(* IEC 61131-3 sources: daoli-st-library/DL_Motion (part 18) *)

(* ---- FB_DL_StackingAlignCtrl.st ---- *)
//==============================================================================
// 功能块：FB_DL_StackingAlignCtrl ｜ 中文名称：叠片对位纠偏控制
// 所属子库：DL_Motion ｜ 版本：v1.0.0 ｜ 兼容：CODESYS V3.5+ / TwinCAT 3 / 汇川 InoProShop
// 功能描述：叠片机 CCD 对位纠偏量的解算件。输入像素偏差与角度偏差，经「像素→机械」
//           标定矩阵的逆映射得机械纠偏量（mm / mrad），输出双轴纠偏指令、超差 NG 与
//           行程限幅标志。标定矩阵求逆委托 FC_DL_Affine2DInvert（组合调用，不复制
//           低层实现）；矩阵奇异时沿用上次有效逆矩阵并置 bMatrixFallback，无历史有效
//           值时判故障。本件只解算纠偏量，不定义轴状态、不发运动指令——轴状态与运动
//           指令的唯一属主是运动层（T1-6 纪律），本件仅输出「允许上层下发纠偏」的
//           bReady 许可位。
// 开源溯源 (Origin)：道莅原创实现（参考 公开工程惯例 分类与参数域）
// 单位表：像素偏差[像素] / 纠偏量[mm] / 角度偏差与角度纠偏量[mrad] / 标定矩阵线性块
//         [mm 每像素] / 标定矩阵平移列[mm] / 行程门限[mm] / 超差门限[mm 或 mrad] /
//         行列式[无量纲]
// 错误码表：16#0004_01EB 信息级（纠偏量被行程限幅，bClamped 置位，限幅后值不得当作
//           正常纠偏量计数，须 HMI 可辨，不置 bError）/ 16#0004_01EC 信息级（标定矩阵
//           退化不可逆，沿用上次有效逆矩阵，bMatrixFallback 置位，不置 bError）/
//           16#0004_030C 故障级（标定矩阵非法/不可逆且无历史有效值，置 bError，纠偏量
//           回零）/ 16#0004_030D 故障级（输入非有限或纠偏解算溢出，置 bError，纠偏量
//           回零）/ 16#0004_030E 故障级兜底（状态机落 ELSE 非法状态，置 bError，纠偏量
//           回零）。码位 16#0004 段，信息带 01xx、故障带 03xx，不越段不挪用预留槽。
// 状态机：E_DL_StackAlignState（eIdle=0 失能/待机 / eAlign=10 正常纠偏解算 /
//           eLimited=20 行程限幅生效 / eCamLost=30 相机无效不纠偏 / eFault=99 故障
//           兜底），CASE 含 ELSE 兜底，ELSE 置 030E 且纠偏量回零 bValid := FALSE。
// 边界行为：① 标定矩阵经 FC_DL_Affine2DInvert 求逆（每拍无条件调用恰好一次）；奇异
//           时若有历史有效逆矩阵 → 信息 01EC + bMatrixFallback := TRUE + 沿用上次值，
//           若无历史有效值 → 故障 030C；② 纠偏量限幅到行程 → bClamped := TRUE +
//           信息 01EB；③ 超差判据取「限幅前」原始纠偏量与角度偏差（限幅会把超差量压成
//           行程端点，用限幅后值判超差会漏判），命中即 bNg := TRUE 并锁存至 bReset；
//           ④ bCamValid := FALSE → 纠偏量回零、bReady := FALSE、bClamped := FALSE、
//           不改 bNg（不做判定即不改判定结果），状态进 eCamLost；⑤ 非有限（NaN 自反判
//           + Inf 幅值上限判，R79）→ 故障 030D 且纠偏量回零；⑥ 失能 → 纠偏量回零 +
//           bReady := FALSE（R72 许可类输出显式 FALSE）；⑦ 行程域倒置（下限 ≥ 上限）
//           按零行程处理，归入 01EB 限幅语义并撤 bReady，不新占码位。
// 修订历史：v1.0.0 2026-11-17 首版（R25 派单 · §4.11，依赖 §4.1 件 FC_DL_Affine2DInvert 语义）
//==============================================================================
(*------------------------------------------------------------------------------
 * 枚举: E_DL_StackAlignState（归属 DL_Motion，与 FB_DL_StackingAlignCtrl 同文件）
 *----------------------------------------------------------------------------*)
TYPE E_DL_StackAlignState :
(
    eIdle    := 0,   // 失能/待机：纠偏量回零，bReady 撤销 / Disabled, corrections zeroed, bReady dropped
    eAlign   := 10,  // 正常解算：纠偏量在行程内，允许上层下发 / Normal solve, corrections within travel
    eLimited := 20,  // 行程限幅生效：纠偏量被夹到行程端点 / Travel clamp active, corrections clipped
    eCamLost := 30,  // 相机无效：不纠偏、不改超差判定 / Camera invalid, no correction, NG untouched
    eFault   := 99   // 故障兜底：矩阵非法/非有限/非法状态 / Fault fallback
);
END_TYPE

(*==============================================================================
 * 功能块: FB_DL_StackingAlignCtrl
 * 调用约定: 每个扫描周期无条件调用一次；像素偏差与角度偏差由上层刷新。
 *============================================================================*)
FUNCTION_BLOCK FB_DL_StackingAlignCtrl
VAR_INPUT
    fOffsetXPx      : LREAL;                       // 像素偏差 X [像素]，正 = 偏右 / Pixel offset X [px], positive = right
    fOffsetYPx      : LREAL;                       // 像素偏差 Y [像素]，正 = 偏下 / Pixel offset Y [px], positive = down
    fAngleMrad      : LREAL;                       // 角度偏差 [mrad]，正 = 逆时针 / Angular offset [mrad], positive = counter-clockwise
    afPixelToMachine : ARRAY[0..2, 0..2] OF LREAL; // 像素→机械标定矩阵 [mm 每像素]，行主序 / Pixel-to-machine calibration matrix [mm per px], row-major
    fAxisXMinMm     : LREAL;                       // 纠偏轴 X 行程下限 [mm] / Correction axis X travel floor [mm]
    fAxisXMaxMm     : LREAL;                       // 纠偏轴 X 行程上限 [mm] / Correction axis X travel ceiling [mm]
    fAxisYMinMm     : LREAL;                       // 纠偏轴 Y 行程下限 [mm] / Correction axis Y travel floor [mm]
    fAxisYMaxMm     : LREAL;                       // 纠偏轴 Y 行程上限 [mm] / Correction axis Y travel ceiling [mm]
    fNgTolMm        : LREAL := 0.05;               // 位置超差门限 [mm] / Position NG tolerance [mm]
    fNgTolMrad      : LREAL := 2.0;                // 角度超差门限 [mrad] / Angular NG tolerance [mrad]
    bCamValid       : BOOL;                        // 相机结果有效（取像成功且特征识别置信） / Camera result valid
    bAxisInPos      : BOOL;                        // 纠偏轴在定位完成状态（上层反馈） / Correction axis in position
    bEnable         : BOOL;                        // 总使能 / Master enable
    bReset          : BOOL;                        // 复位，上升沿清超差锁存与故障 / Reset, rising edge clears NG latch and fault
END_VAR
VAR_OUTPUT
    fCorrXMm        : LREAL;                       // 纠偏量 X [mm]，已按行程限幅 / Correction X [mm], travel-clamped
    fCorrYMm        : LREAL;                       // 纠偏量 Y [mm]，已按行程限幅 / Correction Y [mm], travel-clamped
    fCorrAngleMrad  : LREAL;                       // 角度纠偏量 [mrad] / Angular correction [mrad]
    bNg             : BOOL;                        // 超差判定，锁存至 bReset / Out-of-tolerance latch, cleared by reset
    bClamped        : BOOL;                        // 行程限幅生效标志 / Travel clamp active flag
    bReady          : BOOL;                        // 允许上层下发纠偏（相机有效且在位且在行程内） / Correction may be issued by the upper layer
    bMatrixFallback : BOOL;                        // 沿用上次有效逆矩阵标志 / Reusing the last valid inverse matrix
    eErr            : UDINT;                       // 错误码，0 = 无错，码位 16#0004_01EB 起信息级、16#0004_030C 起故障级（分带见错误码表） / Error code, 0 = no error, band info/fault per the code table
    bError          : BOOL;                        // 故障级标志，仅故障级错误置位 / Fault-class flag, set only on fault-level codes
    bValid          : BOOL;                        // 纠偏量可用标志，失能/故障闸显式 FALSE / Correction usable flag, explicit FALSE on disable/fault gates
    eState          : E_DL_StackAlignState;        // 主状态机当前状态 / Current state of the main state machine
END_VAR
VAR
    fbReset         : R_TRIG;                      // 复位上升沿检测实例 / Reset rising edge detector
    afMInvNew       : ARRAY[0..2, 0..2] OF LREAL;  // 本拍求得的逆矩阵 [mm 每像素] / Inverse matrix of this scan
    afMInvLast      : ARRAY[0..2, 0..2] OF LREAL;  // 上次有效逆矩阵（退化时沿用）[mm 每像素] / Last valid inverse matrix
    afMInvEff       : ARRAY[0..2, 0..2] OF LREAL;  // 本拍生效逆矩阵（新值或沿用值）[mm 每像素] / Effective inverse matrix of this scan
    nI              : INT;                         // 行循环索引 [—] / Row loop index
    nJ              : INT;                         // 列循环索引 [—] / Column loop index
    uInvErr         : UDINT;                       // 求逆件错误码暂存 / Inverse-function error code staging
    fDetNew         : LREAL;                       // 本拍线性块行列式 [无量纲] / Linear block determinant of this scan
    bInvFault       : BOOL;                        // 求逆件故障标志暂存 / Inverse-function fault flag staging
    bInvValid       : BOOL;                        // 求逆件结果可用暂存 / Inverse-function usable flag staging
    bInvOk          : BOOL;                        // 求逆件返回值暂存（与可用标志同口径） / Inverse-function return staging
    bHasValidInv    : BOOL;                        // 已存在历史有效逆矩阵 / A valid inverse matrix has been stored
    fRawXMm         : LREAL;                       // 限幅前纠偏量 X [mm] / Unclamped correction X [mm]
    fRawYMm         : LREAL;                       // 限幅前纠偏量 Y [mm] / Unclamped correction Y [mm]
    fLimX           : LREAL;                       // 生效 X 行程上限（倒置时夹零）[mm] / Effective X travel ceiling [mm]
    fLimY           : LREAL;                       // 生效 Y 行程上限（倒置时夹零）[mm] / Effective Y travel ceiling [mm]
    bTravelXBad     : BOOL;                        // X 行程域倒置标志 / X travel range inverted flag
    bTravelYBad     : BOOL;                        // Y 行程域倒置标志 / Y travel range inverted flag
    bNonFin         : BOOL;                        // 非有限判定中间标志 / Non-finite detection intermediate flag
    bFirstScan      : BOOL := TRUE;                // 上电首拍标志 / First-scan flag
END_VAR
VAR CONSTANT
    DL_SAC_CODE_INFO_1 : UDINT := 16#0004_01EB;    // 信息级槽 1（纠偏量被行程限幅） / info slot 1
    DL_SAC_CODE_INFO_2 : UDINT := 16#0004_01EC;    // 信息级槽 2（标定矩阵退化沿用上次） / info slot 2
    DL_SAC_CODE_FLT_1  : UDINT := 16#0004_030C;    // 故障级槽 1（矩阵非法且无历史有效值） / fault slot 1
    DL_SAC_CODE_FLT_2  : UDINT := 16#0004_030D;    // 故障级槽 2（输入非有限/解算溢出） / fault slot 2
    DL_SAC_CODE_FLT_3  : UDINT := 16#0004_030E;    // 故障级槽 3（非法状态兜底） / fault slot 3, illegal-state fallback
    DL_SAC_DET_EPS     : LREAL := 1.0E-9;          // 逆矩阵相对奇异判据 [无量纲] / Relative singularity threshold of the inverse
    DL_SAC_ZERO        : LREAL := 0.0;             // 零值常量，避免裸字面量 [—] / Zero constant, avoids a bare literal
    DL_SAC_TOL         : LREAL := 1.0E-6;          // 浮点比较容差 [—] / Float comparison tolerance
    DL_SAC_INF         : LREAL := 1.7976931348623157E308; // LREAL 幅值上限，Inf 判据 / LREAL magnitude ceiling, Inf criterion
END_VAR

(*------------------------------------------------------------------------------
 * 段 1｜无条件刷新区（红线 5）：复位沿检测在任何分支之外周期调用
 *----------------------------------------------------------------------------*)
fbReset(CLK := bReset);                            // 复位沿检测无条件刷新 / reset edge refreshed unconditionally

(*------------------------------------------------------------------------------
 * 段 2｜复位沿处理（改写置于沿后，防吞沿 R39）：清超差锁存与故障码；
 *       历史有效逆矩阵属标定事实，不随复位清除（头注释边界行为①）
 *----------------------------------------------------------------------------*)
IF fbReset.Q THEN
    bNg     := FALSE;                              // 超差锁存清除 / NG latch cleared
    bError  := FALSE;                              // 故障标志清除 / fault flag cleared
    eErr    := 16#0000_0000;                       // 错误码清除 / error code cleared
    eState  := E_DL_StackAlignState.eIdle;         // 回待机 / back to idle
    bFirstScan := TRUE;                            // 重新首拍化 / re-initialize first scan
END_IF

(*------------------------------------------------------------------------------
 * 段 3｜非有限输入闸（标量、行程、门限逐个：NaN 自反判 + Inf 幅值上限判）
 *       命中即纠偏量回零 + 撤许可，安全侧不留上次值（红线 6）
 *----------------------------------------------------------------------------*)
bNonFin := (fOffsetXPx <> fOffsetXPx) OR (ABS(fOffsetXPx) >= DL_SAC_INF)
        OR (fOffsetYPx <> fOffsetYPx) OR (ABS(fOffsetYPx) >= DL_SAC_INF)
        OR (fAngleMrad <> fAngleMrad) OR (ABS(fAngleMrad) >= DL_SAC_INF)
        OR (fAxisXMinMm <> fAxisXMinMm) OR (ABS(fAxisXMinMm) >= DL_SAC_INF)
        OR (fAxisXMaxMm <> fAxisXMaxMm) OR (ABS(fAxisXMaxMm) >= DL_SAC_INF)
        OR (fAxisYMinMm <> fAxisYMinMm) OR (ABS(fAxisYMinMm) >= DL_SAC_INF)
        OR (fAxisYMaxMm <> fAxisYMaxMm) OR (ABS(fAxisYMaxMm) >= DL_SAC_INF)
        OR (fNgTolMm <> fNgTolMm) OR (ABS(fNgTolMm) >= DL_SAC_INF)
        OR (fNgTolMrad <> fNgTolMrad) OR (ABS(fNgTolMrad) >= DL_SAC_INF); // 引脚非有限汇总判定 / aggregated non-finite check
IF bNonFin THEN
    eState := E_DL_StackAlignState.eFault;          // 进故障相 / enter fault state
    eErr   := DL_SAC_CODE_FLT_2;                    // 故障级：输入非有限 / fault: non-finite input
    bError := TRUE;                                 // 故障级必置 bError（R45 配对）/ fault-class pairs with bError
    bValid := FALSE;                                // 输出不可用 / outputs unusable
    fCorrXMm := DL_SAC_ZERO;                        // 纠偏量回零安全侧 / correction zeroed, safe side
    fCorrYMm := DL_SAC_ZERO;                        // 纠偏量回零安全侧 / correction zeroed, safe side
    fCorrAngleMrad := DL_SAC_ZERO;                  // 角度纠偏回零安全侧 / angular correction zeroed
    bClamped := FALSE;                              // 限幅标志撤 / clamp flag withdrawn
    bReady := FALSE;                                // 许可撤（R72）/ permission dropped
    bMatrixFallback := FALSE;                       // 降级标志撤 / fallback flag withdrawn
    RETURN;
END_IF

(*------------------------------------------------------------------------------
 * 段 4｜标定矩阵求逆：组合调用 FC_DL_Affine2DInvert（每拍无条件调用恰好一次，
 *       禁止复制低层 2x2 伴随求逆实现）；引脚契约以源码头注释为准
 *----------------------------------------------------------------------------*)
bInvOk := FC_DL_Affine2DInvert(afM := afPixelToMachine,   // 待求逆标定矩阵 [mm 每像素] / calibration matrix to invert
                               fDetEps := DL_SAC_DET_EPS, // 相对奇异判据 [无量纲] / relative singularity threshold
                               afMInv => afMInvNew,       // 逆矩阵输出 [mm 每像素] / inverse matrix output
                               fDet => fDetNew,           // 行列式输出 [无量纲] / determinant output
                               eErr => uInvErr,           // 下游错误码暂存 / downstream error code staging
                               bError => bInvFault,       // 下游故障标志暂存 / downstream fault flag staging
                               bValid => bInvValid);      // 下游可用标志暂存 / downstream usable flag staging

(*------------------------------------------------------------------------------
 * 段 5｜逆矩阵不可用降级：有历史有效值 → 信息 01EC 沿用上次；无历史 → 故障 030C。
 *       下游信息级码不升格为故障（§5.5 纪律），仅在逆结果不可用时按本件语义处置
 *----------------------------------------------------------------------------*)
IF (NOT bInvValid) OR (NOT bInvOk) THEN
    IF bHasValidInv THEN
        FOR nI := 0 TO 2 DO
            FOR nJ := 0 TO 2 DO
                afMInvEff[nI, nJ] := afMInvLast[nI, nJ];   // 沿用上次有效逆矩阵 / reuse the last valid inverse
            END_FOR
        END_FOR
        bMatrixFallback := TRUE;                   // 降级标志置位 / fallback flag raised
        eState := E_DL_StackAlignState.eAlign;     // 按正常解算相继续 / continue in the normal solve state
        eErr   := DL_SAC_CODE_INFO_2;              // 信息级：矩阵退化沿用上次（不置 bError）/ info: singular matrix, last valid reused
        bError := FALSE;                           // 信息级不置 bError（R45/R101）/ info never raises bError
    ELSE
        eState := E_DL_StackAlignState.eFault;     // 进故障相 / enter fault state
        eErr   := DL_SAC_CODE_FLT_1;               // 故障级：矩阵非法且无历史有效值 / fault: illegal matrix with no history
        bError := TRUE;                            // 故障级必置 bError（R45 配对）/ fault-class pairs with bError
        bValid := FALSE;                           // 输出不可用 / outputs unusable
        fCorrXMm := DL_SAC_ZERO;                   // 纠偏量回零安全侧 / correction zeroed, safe side
        fCorrYMm := DL_SAC_ZERO;                   // 纠偏量回零安全侧 / correction zeroed, safe side
        fCorrAngleMrad := DL_SAC_ZERO;             // 角度纠偏回零安全侧 / angular correction zeroed
        bClamped := FALSE;                         // 限幅标志撤 / clamp flag withdrawn
        bReady := FALSE;                           // 许可撤（R72）/ permission dropped
        bMatrixFallback := FALSE;                  // 无历史可沿用，降级标志不得冒充 / fallback flag must not fake reuse
        RETURN;
    END_IF
ELSE
    FOR nI := 0 TO 2 DO
        FOR nJ := 0 TO 2 DO
            afMInvEff[nI, nJ] := afMInvNew[nI, nJ];        // 采用本拍逆矩阵 / take the inverse of this scan
            afMInvLast[nI, nJ] := afMInvNew[nI, nJ];       // 记账：历史有效逆矩阵 / bookkeeping: last valid inverse
        END_FOR
    END_FOR
    bHasValidInv := TRUE;                          // 历史有效值成立 / history becomes valid
    bMatrixFallback := FALSE;                      // 正常路径不置降级 / no fallback on the normal path
END_IF

(*------------------------------------------------------------------------------
 * 段 6｜相机无效闸：不纠偏、撤许可、不改超差判定（两条退出条件在 CASE eCamLost 相）
 *----------------------------------------------------------------------------*)
IF NOT bCamValid THEN
    fCorrXMm := DL_SAC_ZERO;                       // 纠偏量回零（不纠偏）/ correction zeroed, no correction
    fCorrYMm := DL_SAC_ZERO;                       // 纠偏量回零（不纠偏）/ correction zeroed, no correction
    fCorrAngleMrad := DL_SAC_ZERO;                 // 角度纠偏回零 / angular correction zeroed
    bClamped := FALSE;                             // 限幅标志撤 / clamp flag withdrawn
    bReady := FALSE;                               // 许可撤（R72）/ permission dropped
    bValid := FALSE;                               // 纠偏量不可用 / corrections unusable
    eErr   := 16#0000_0000;                        // 相机无效不占码位（无对应分配槽）/ no code allocated for a camera dropout
    bError := FALSE;                               // 不升格为故障 / not escalated to a fault
    IF bEnable THEN
        eState := E_DL_StackAlignState.eCamLost;   // 相机丢失相 / camera-lost state
    ELSE
        eState := E_DL_StackAlignState.eIdle;      // 失能优先回待机 / disable outranks, back to idle
    END_IF
    // 超差锁存原样保持：本拍不做判定即不改判定结果，绝不在此处清 bNg / NG latch held verbatim, never cleared here
    RETURN;
END_IF

(*------------------------------------------------------------------------------
 * 段 7｜纠偏量解算：逆映射 p_mech = M^(-1) x [dx_px, dy_px, 1]^T，
 *       角度纠偏量按标定链直通（本件不另设角度增益，增益归标定矩阵）
 *----------------------------------------------------------------------------*)
fRawXMm := afMInvEff[0, 0] * fOffsetXPx + afMInvEff[0, 1] * fOffsetYPx + afMInvEff[0, 2];   // 纠偏量 X [mm] / correction X [mm]
fRawYMm := afMInvEff[1, 0] * fOffsetXPx + afMInvEff[1, 1] * fOffsetYPx + afMInvEff[1, 2];   // 纠偏量 Y [mm] / correction Y [mm]
fCorrAngleMrad := fAngleMrad;                      // 角度纠偏量直通 [mrad] / angular correction passed through
IF (fRawXMm <> fRawXMm) OR (ABS(fRawXMm) >= DL_SAC_INF)
   OR (fRawYMm <> fRawYMm) OR (ABS(fRawYMm) >= DL_SAC_INF) THEN
    eState := E_DL_StackAlignState.eFault;         // 解算溢出进故障相 / solve overflow enters fault state
    eErr   := DL_SAC_CODE_FLT_2;                   // 故障级：解算结果非有限（复用输入非法槽）/ fault: non-finite result, shares the input slot
    bError := TRUE;                                // 故障级必置 bError（R45 配对）/ fault-class pairs with bError
    bValid := FALSE;                               // 输出不可用 / outputs unusable
    fCorrXMm := DL_SAC_ZERO;                       // 纠偏量回零安全侧 / correction zeroed, safe side
    fCorrYMm := DL_SAC_ZERO;                       // 纠偏量回零安全侧 / correction zeroed, safe side
    fCorrAngleMrad := DL_SAC_ZERO;                 // 角度纠偏回零安全侧 / angular correction zeroed
    bClamped := FALSE;                             // 限幅标志撤 / clamp flag withdrawn
    bReady := FALSE;                               // 许可撤（R72）/ permission dropped
    RETURN;
END_IF

(*------------------------------------------------------------------------------
 * 段 8｜行程限幅：先判行程域（下限 ≥ 上限 → 零行程），再逐轴夹取；
 *       一旦夹取即置 bClamped + 信息 01EB（限幅值不得当正常纠偏量计数）
 *----------------------------------------------------------------------------*)
bTravelXBad := (fAxisXMinMm >= fAxisXMaxMm - DL_SAC_TOL);   // X 行程域倒置判定 / X travel inverted predicate
bTravelYBad := (fAxisYMinMm >= fAxisYMaxMm - DL_SAC_TOL);   // Y 行程域倒置判定 / Y travel inverted predicate
IF bTravelXBad THEN
    fLimX := fAxisXMinMm;                          // 零行程：上限夹到下限 / zero travel: ceiling pinned to the floor
ELSE
    fLimX := fAxisXMaxMm;                          // 正常行程上限 / normal travel ceiling
END_IF
IF bTravelYBad THEN
    fLimY := fAxisYMinMm;                          // 零行程：上限夹到下限 / zero travel: ceiling pinned to the floor
ELSE
    fLimY := fAxisYMaxMm;                          // 正常行程上限 / normal travel ceiling
END_IF
bClamped := FALSE;                                 // 限幅标志逐拍重判 / clamp flag re-judged per scan
fCorrXMm := fRawXMm;                               // 先取原始值再夹取 / take the raw value before clipping
IF fCorrXMm > fLimX THEN
    fCorrXMm := fLimX;                             // 上限夹取 [mm] / clipped to the ceiling
    bClamped := TRUE;                              // 限幅生效 / clamp active
END_IF
IF fCorrXMm < fAxisXMinMm THEN
    fCorrXMm := fAxisXMinMm;                       // 下限夹取 [mm] / clipped to the floor
    bClamped := TRUE;                              // 限幅生效 / clamp active
END_IF
fCorrYMm := fRawYMm;                               // 先取原始值再夹取 / take the raw value before clipping
IF fCorrYMm > fLimY THEN
    fCorrYMm := fLimY;                             // 上限夹取 [mm] / clipped to the ceiling
    bClamped := TRUE;                              // 限幅生效 / clamp active
END_IF
IF fCorrYMm < fAxisYMinMm THEN
    fCorrYMm := fAxisYMinMm;                       // 下限夹取 [mm] / clipped to the floor
    bClamped := TRUE;                              // 限幅生效 / clamp active
END_IF

(*------------------------------------------------------------------------------
 * 段 9｜超差判定与锁存：判据取限幅前原始量（限幅后值被压成行程端点会漏判超差），
 *       命中即锁存 bNg，仅 bReset 可清（超差件不因下一拍合格而自动放行）
 *----------------------------------------------------------------------------*)
IF (ABS(fRawXMm) > fNgTolMm) OR (ABS(fRawYMm) > fNgTolMm)
   OR (ABS(fCorrAngleMrad) > fNgTolMrad) THEN
    bNg := TRUE;                                   // 超差锁存 / NG latched
END_IF

(*------------------------------------------------------------------------------
 * 段 10｜状态机：CASE 含 ELSE 兜底（非法状态 → 030E + 纠偏量回零 + 撤许可）
 *        eCamLost 与 eFault 相各给两条以上退出条件（事件沿之外必含前置消失）
 *----------------------------------------------------------------------------*)
CASE eState OF

    E_DL_StackAlignState.eIdle:
        bValid := FALSE;                           // 失能闸显式不可用（R72）/ explicit FALSE on the disable gate
        bReady := FALSE;                           // 许可撤 / permission dropped
        fCorrXMm := DL_SAC_ZERO;                   // 纠偏量回零安全侧 / correction zeroed, safe side
        fCorrYMm := DL_SAC_ZERO;                   // 纠偏量回零安全侧 / correction zeroed, safe side
        fCorrAngleMrad := DL_SAC_ZERO;             // 角度纠偏回零安全侧 / angular correction zeroed
        bClamped := FALSE;                         // 限幅标志撤 / clamp flag withdrawn
        bMatrixFallback := FALSE;                  // 降级标志撤 / fallback flag withdrawn
        eErr := 16#0000_0000;                      // 待机无错 / no error in idle
        bError := FALSE;                           // 待机无故障 / no fault in idle
        IF bEnable AND bCamValid THEN
            eState := E_DL_StackAlignState.eAlign; // 使能且相机有效进解算相 / enable with a valid camera enters solve
            bFirstScan := FALSE;                   // 首拍标志清除 / first-scan flag cleared
        END_IF

    E_DL_StackAlignState.eAlign:
        bValid := TRUE;                            // 纠偏量可用 / corrections usable
        bError := FALSE;                           // 解算相无故障 / no fault in the solve state
        IF bClamped THEN
            eErr := DL_SAC_CODE_INFO_1;            // 信息级：限幅生效 / info: clamp active
            eState := E_DL_StackAlignState.eLimited;   // 转限幅相 / enter the limited state
        ELSE
            eErr := 16#0000_0000;                  // 行程内无错 / within travel, no error
        END_IF
        bReady := bAxisInPos AND bCamValid;        // 在位且相机有效才允许下发 / issue only when in position and camera valid
        IF NOT bEnable THEN
            eState := E_DL_StackAlignState.eIdle;  // 失能回待机 / disable returns to idle
            bValid := FALSE;                       // 失能闸显式不可用 / explicit FALSE on the disable gate
            bReady := FALSE;                       // 许可撤 / permission dropped
        ELSIF NOT bCamValid THEN
            eState := E_DL_StackAlignState.eCamLost;   // 相机丢失转丢失相 / camera dropout enters the lost state
            bValid := FALSE;                       // 输出不可用 / outputs unusable
            bReady := FALSE;                       // 许可撤 / permission dropped
        END_IF

    E_DL_StackAlignState.eLimited:
        bValid := TRUE;                            // 限幅后值可用（须 HMI 可辨）/ clipped values usable, flagged for HMI
        bError := FALSE;                           // 信息级不置 bError / info never raises bError
        eErr := DL_SAC_CODE_INFO_1;                // 信息级：纠偏量被行程限幅 / info: correction clamped by travel
        bReady := bAxisInPos AND bCamValid AND (NOT bTravelXBad) AND (NOT bTravelYBad);   // 行程域倒置时撤许可 / travel range inverted drops permission
        IF NOT bEnable THEN
            eState := E_DL_StackAlignState.eIdle;  // 失能回待机（退出条件一）/ disable returns to idle, first exit
            bValid := FALSE;                       // 失能闸显式不可用 / explicit FALSE on the disable gate
            bReady := FALSE;                       // 许可撤 / permission dropped
        ELSIF NOT bCamValid THEN
            eState := E_DL_StackAlignState.eCamLost;   // 相机丢失（退出条件二）/ camera dropout, second exit
            bValid := FALSE;                       // 输出不可用 / outputs unusable
            bReady := FALSE;                       // 许可撤 / permission dropped
        ELSIF NOT bClamped THEN
            eState := E_DL_StackAlignState.eAlign; // 限幅消失回解算相（退出条件三）/ clamp gone, third exit to solve
        END_IF

    E_DL_StackAlignState.eCamLost:
        bValid := FALSE;                           // 输出不可用 / outputs unusable
        bReady := FALSE;                           // 许可撤 / permission dropped
        fCorrXMm := DL_SAC_ZERO;                   // 纠偏量回零安全侧 / correction zeroed, safe side
        fCorrYMm := DL_SAC_ZERO;                   // 纠偏量回零安全侧 / correction zeroed, safe side
        fCorrAngleMrad := DL_SAC_ZERO;             // 角度纠偏回零安全侧 / angular correction zeroed
        bClamped := FALSE;                         // 限幅标志撤 / clamp flag withdrawn
        eErr := 16#0000_0000;                      // 相机丢失不占码位 / no code allocated for a camera dropout
        bError := FALSE;                           // 不升格为故障 / not escalated to a fault
        IF bEnable AND bCamValid THEN
            eState := E_DL_StackAlignState.eAlign; // 相机恢复且使能回解算相（退出条件一）/ camera back, first exit
        ELSIF NOT bEnable THEN
            eState := E_DL_StackAlignState.eIdle;  // 失能回待机（退出条件二）/ disable, second exit
        END_IF

    E_DL_StackAlignState.eFault:
        bValid := FALSE;                           // 故障闸显式不可用（R72）/ explicit FALSE on the fault gate
        bReady := FALSE;                           // 许可撤 / permission dropped
        fCorrXMm := DL_SAC_ZERO;                   // 纠偏量回零安全侧 / correction zeroed, safe side
        fCorrYMm := DL_SAC_ZERO;                   // 纠偏量回零安全侧 / correction zeroed, safe side
        fCorrAngleMrad := DL_SAC_ZERO;             // 角度纠偏回零安全侧 / angular correction zeroed
        bClamped := FALSE;                         // 限幅标志撤 / clamp flag withdrawn
        IF eErr = 16#0000_0000 THEN
            eErr := DL_SAC_CODE_FLT_1;             // 入口无码时按矩阵非法解释（R45：bError 必须有对应码）/ default to the matrix slot so bError always maps to a code
        END_IF
        bError := TRUE;                            // 故障级必置 bError（R45 配对）/ fault-class pairs with bError
        IF bEnable AND bInvValid AND bCamValid AND bHasValidInv THEN
            eState := E_DL_StackAlignState.eAlign; // 前置条件全部恢复才回解算相（退出条件 ≥2）/ only when every precondition recovers
        END_IF

    ELSE
        eState := E_DL_StackAlignState.eFault;     // 非法状态兜底 / illegal-state fallback
        eErr := DL_SAC_CODE_FLT_3;                 // 故障级兜底：非法状态 / fault fallback: illegal state
        bError := TRUE;                            // 故障级必置 bError（R45 配对）/ fault-class pairs with bError
        bValid := FALSE;                           // 输出不可用 / outputs unusable
        bReady := FALSE;                           // 许可撤 / permission dropped
        fCorrXMm := DL_SAC_ZERO;                   // 纠偏量回零安全侧 / correction zeroed, safe side
        fCorrYMm := DL_SAC_ZERO;                   // 纠偏量回零安全侧 / correction zeroed, safe side
        fCorrAngleMrad := DL_SAC_ZERO;             // 角度纠偏回零安全侧 / angular correction zeroed

END_CASE
END_FUNCTION_BLOCK

(* ---- FB_DL_StepperFeederBelt.st ---- *)
(*==============================================================================
 * 组件名称 (Component)  : FB_DL_StepperFeederBelt
 * 所属子库 (Sublibrary) : DL_Motion
 * 当前版本 (Version)    : 1.0.0
 * 兼容性 (Platform)     : CODESYS 3.5 / TwinCAT 3 / 汇川 InoProShop（纯标准元素，零方言）
 * 功能描述 (Function)   : 步进供料带间歇送料 + 色标偏差补偿。送料请求上升沿受理一次，
 *                         步距 = 标称间距 + 色标补偿增量（偏差 × 增益），补偿量按上限
 *                         累计约束；送料后等停稳确认时长再给单拍完成脉冲。运行期请求
 *                         一律丢弃不排队。不做色标检测本身（偏差由引脚注入）、不做
 *                         速度前馈、不做多段送料。
 *                         说明：接口契约 MoveRelative 只接受距离与速度，fAccel_mmS2 仅参与
 *                         参数门禁校验，不向下转发（规格口径在本行登记）。
 * 溯源 (Origin)         : 道莅 clean-room 防御性实现
 * 本文件内含 (Contains) : TYPE E_DL_FeederState / FUNCTION_BLOCK FB_DL_StepperFeederBelt
 * 依赖 (Depends)        : DL_Device/I_DL_StepperOpenLoop（只调用契约方法与属性）
 * 红线自检 (Redline)    : 无外部全局变量、无硬件地址直引 ｜ 全变量中英双语同行注释
 *                         间距判零防除零 ｜ 步距双向钳制（防倒料） ｜ 非有限用自反比较
 *                         枚举显式赋值 ｜ 停稳定时器与沿检测无条件周期刷新 ｜ CASE 含 ELSE
 * 错误码表 (Codes)      : 16#0004_032C 就绪/单次送料完成
 *                         16#0004_032D 故障级 步进轴拒绝送料指令。反证句：轴拒绝在输出侧
 *                                    与「组态非法」同为「本拍无位移」，但组态非法可由 032E
 *                                    在启动前观测，故轴拒绝须独立成码
 *                         16#0004_032E 故障级 组态非法（间距判零、增益/上限/速度/加速度出域）
 *                         16#0004_032F 信息级 补偿后步距越 0.5~1.5 倍间距已钳制（防倒料，
 *                                    不置故障级标志，送料照常进行）
 *                         16#0004_0330 故障级 累计补偿越上限，停送（继续补偿会把误差藏进
 *                                    机构行程）。本件 5 槽全用、无预留槽，已登记待裁定
 * 修订历史 (Revision)   : 2026-11-17  v1.0.0  首版入库 · R28 · 阶段三批 1
 * 验收向量 (Acceptance) : 正向 间距 100 mm、偏差 +2 mm、增益 0.5 → 步距 101 mm、累计
 *                         +1 mm、16#0004_032C、计数 +1
 *                         反向 连续 60 拍偏差 +1 mm（增益 0.5）→ 累计 30 mm 超上限 20 mm
 *                         → 16#0004_0330 停送；间距给 0 → 16#0004_032E；步距被钳到
 *                         1.5 倍间距 → 16#0004_032F 且照常送料
 *============================================================================*)

(*-----------------------------------------------------------------------------
 * 枚举: E_DL_FeederState（归属本功能块，同文件发布，全库唯一定义）
 * 含义: 供料带送料相位，每个成员在 CASE 中有且仅有一个标签。
 *----------------------------------------------------------------------------*)
TYPE E_DL_FeederState :
(
    eIdle     := 0,    // 空闲：等送料请求沿 / Idle, waiting for the index request edge
    eIndexing := 10,   // 送料中：已派单，等轴就绪 / Indexing, dispatched and waiting for the axis to be ready
    eSettling := 20,   // 停稳确认：等 tSettle 计时满 / Settling, waiting for the settle time
    eFault    := 99    // 故障：锁存码保持，仅使能沿重启 / Fault, the latch code is held until an enable edge
);
END_TYPE

FUNCTION_BLOCK FB_DL_StepperFeederBelt
VAR_INPUT
    bEnable         : BOOL := FALSE;      // 使能，上升沿清补偿累计（班次重启语义） / Enable, the rising edge clears the trim accumulation
    bIndexReq       : BOOL := FALSE;      // 送料请求，上升沿受理，运行期丢弃 / Index request, accepted on the rising edge and dropped while busy
    fPitch_mm       : REAL := 100.0;      // 标称间距 [mm]，域 1~2000 / Nominal pitch in millimetres, domain 1 to 2000
    fMarkOffset_mm  : REAL := 0.0;        // 色标偏差 [mm]，域 ±20，正=超前 / Mark offset in millimetres, domain plus minus 20, positive means ahead
    fTrimGain       : REAL := 0.5;        // 补偿增益 [—]，域 0~1（>1 振荡） / Trim gain, domain 0 to 1, above 1 oscillates
    fTrimAccumMax_mm : REAL := 20.0;      // 累计补偿上限 [mm]，域 0.5~50 / Trim accumulation limit in millimetres, domain 0.5 to 50
    fSpeed_mmS      : REAL := 100.0;      // 运行速度 [mm/s]，域 1~500 / Run speed in millimetres per second, domain 1 to 500
    fAccel_mmS2     : REAL := 1000.0;     // 加速度 [mm/s²]，域 10~5000（仅门禁校验） / Acceleration, domain 10 to 5000, gate check only
    tSettle         : TIME := T#200MS;    // 停稳确认时长 [ms]，域 10~500 / Settle confirmation time, domain 10 to 500 ms
END_VAR
VAR_IN_OUT
    iAxis           : I_DL_StepperOpenLoop; // 供料带开环步进契约引用 [—] / Feeder belt open-loop stepper contract reference
END_VAR
VAR_OUTPUT
    fStepCmd_mm     : REAL;               // 本次实际步距（含补偿）[mm] / Effective step distance including trim
    fTrimAccum_mm   : REAL;               // 累计补偿量 [mm] / Accumulated trim in millimetres
    bDone           : BOOL;               // 送料完成脉冲，单拍有效 / Index completion pulse, valid for one scan
    bBusy           : BOOL;               // 送料进行中 / Index in progress
    bError          : BOOL;               // 故障级标志，仅故障级码置位 / Fault-class flag, set on fault codes only
    uIndexCnt       : UDINT;              // 累计送料次数 [次] / Total index count
    eErr            : UDINT;              // 错误码，段位 16#0004_xxxx / Error code in segment 16#0004_xxxx
END_VAR
VAR
    _eState         : E_DL_FeederState := E_DL_FeederState.eIdle; // 当前相位 / Current phase
    _bInit          : BOOL := FALSE;      // 首扫标志，取非判定 / First-scan flag, tested negated
    _bRefOk         : BOOL;               // 契约引用有效标志 / Contract reference valid flag
    _bParamOk       : BOOL;               // 参数门禁通过标志 / Parameter gate pass flag
    _bIssueScan     : BOOL;               // 派单当拍标志（本拍不判就绪） / Dispatch scan flag, readiness is not judged in this scan
    _bFaultLatch    : BOOL;               // 故障锁存标志 / Fault latch flag
    _fStepRaw       : REAL;               // 补偿后原始步距 [mm] / Raw step distance after trim
    _fStepEff       : REAL;               // 钳制后生效步距 [mm] / Effective step distance after clamping
    _fAccumNew      : REAL;               // 拟施加的累计补偿 [mm] / Trim accumulation to be applied
    _fSpeedEff      : REAL := 100.0;      // 生效速度（下限兜底）[mm/s] / Effective speed with a lower bound guard
    _uLatchCode     : UDINT;              // 锁存码载体 / Latch code carrier
    _rtrigIndex     : R_TRIG;             // 送料请求上升沿 / Rising edge of the index request
    _rtrigEnable    : R_TRIG;             // 使能上升沿 / Rising edge of the enable input
    _tonSettle      : TON;                // 停稳确认计时 / Settle confirmation timer
END_VAR
VAR CONSTANT
    DL_FDR_READY      : UDINT := 16#0004_032C;  // 就绪/完成码 / Ready or completion code
    DL_FDR_AXIS_REJ   : UDINT := 16#0004_032D;  // 故障级轴拒绝码 / Fault code for a rejected axis command
    DL_FDR_CFG_BAD    : UDINT := 16#0004_032E;  // 故障级组态非法码 / Fault code for bad configuration
    DL_FDR_CLAMP      : UDINT := 16#0004_032F;  // 信息级步距钳制码 / Info code for a clamped step distance
    DL_FDR_ACCUM_MAX  : UDINT := 16#0004_0330;  // 故障级累计补偿越限码 / Fault code for trim accumulation overflow
    DL_FDR_PITCH_LO   : REAL := 1.0;            // 间距下限 [mm] / Pitch lower bound
    DL_FDR_PITCH_HI   : REAL := 2000.0;         // 间距上限 [mm] / Pitch upper bound
    DL_FDR_OFF_HI     : REAL := 20.0;           // 色标偏差绝对值上限 [mm] / Absolute mark offset bound
    DL_FDR_GAIN_HI    : REAL := 1.0;            // 补偿增益上限 [—] / Trim gain upper bound
    DL_FDR_ACCUM_LO   : REAL := 0.5;            // 累计上限下限 [mm] / Lower bound of the accumulation limit
    DL_FDR_ACCUM_HI   : REAL := 50.0;           // 累计上限上限 [mm] / Upper bound of the accumulation limit
    DL_FDR_SPD_LO     : REAL := 1.0;            // 速度下限 [mm/s] / Speed lower bound
    DL_FDR_SPD_HI     : REAL := 500.0;          // 速度上限 [mm/s] / Speed upper bound
    DL_FDR_STEP_LO_K  : REAL := 0.5;            // 步距下限系数 [倍间距] / Step distance lower factor
    DL_FDR_STEP_HI_K  : REAL := 1.5;            // 步距上限系数 [倍间距] / Step distance upper factor
    DL_FDR_EPS        : REAL := 1.0E-6;         // 浮点判零容差 [—] / Float zero tolerance
END_VAR

// 段 1｜输出与单拍标志预置
bDone := FALSE;                                     // 完成脉冲预清 / Completion pulse pre-cleared
bBusy := FALSE;                                     // 运行标志预清 / Busy flag pre-cleared
bError := FALSE;                                    // 故障标志预清 / Fault flag pre-cleared
eErr := 0;                                          // 错误码预清 / Error code pre-cleared
_bIssueScan := FALSE;                               // 派单当拍标志预清 / Dispatch scan flag pre-cleared

// 段 2｜沿检测无条件周期刷新（严禁置于分支内）
_rtrigIndex(CLK := bIndexReq);                      // 送料请求沿 / Index request edge
_rtrigEnable(CLK := bEnable);                       // 使能沿 / Enable edge

// 段 2.5｜停稳定时器无条件周期刷新（仅在停稳相计时）
_tonSettle(IN := (_eState = E_DL_FeederState.eSettling), PT := tSettle);

// 段 3｜首扫初始化（判据取非，R19）
IF NOT _bInit THEN
    _eState := E_DL_FeederState.eIdle;              // 相位待机起步 / Phase starts idle
    _bInit := TRUE;                                 // 首扫只做一次 / The first scan runs once
END_IF

// 段 4｜使能上升沿：清补偿累计与锁存（班次重启语义）
IF _rtrigEnable.Q THEN
    _bFaultLatch := FALSE;                          // 使能沿为锁存解除路径 / The enable edge releases the latch
    _uLatchCode := 0;                               // 锁存码清 / Latch code cleared
    _fAccumNew := 0.0;                              // 累计补偿清零（班次重启）[mm] / Trim accumulation cleared at shift restart
    _eState := E_DL_FeederState.eIdle;              // 相位复位 / Phase reset
END_IF

// 段 5｜契约引用有效性 + 参数门禁逐拍重算（非有限用自反比较）
_bRefOk := (iAxis <> 0);                            // 引用注入判据 / Reference injected flag
_bParamOk := _bRefOk
         AND NOT ((fPitch_mm <> fPitch_mm) OR ((fPitch_mm - fPitch_mm) <> (fPitch_mm - fPitch_mm)))
         AND NOT ((fMarkOffset_mm <> fMarkOffset_mm) OR ((fMarkOffset_mm - fMarkOffset_mm) <> (fMarkOffset_mm - fMarkOffset_mm)))
         AND NOT ((fTrimGain <> fTrimGain) OR ((fTrimGain - fTrimGain) <> (fTrimGain - fTrimGain)))
         AND NOT ((fTrimAccumMax_mm <> fTrimAccumMax_mm) OR ((fTrimAccumMax_mm - fTrimAccumMax_mm) <> (fTrimAccumMax_mm - fTrimAccumMax_mm)))
         AND (fPitch_mm >= DL_FDR_PITCH_LO) AND (fPitch_mm <= DL_FDR_PITCH_HI)
         AND (ABS(fMarkOffset_mm) <= DL_FDR_OFF_HI)
         AND (fTrimGain >= 0.0) AND (fTrimGain <= DL_FDR_GAIN_HI)
         AND (fTrimAccumMax_mm >= DL_FDR_ACCUM_LO) AND (fTrimAccumMax_mm <= DL_FDR_ACCUM_HI)
         AND (fSpeed_mmS >= DL_FDR_SPD_LO) AND (fSpeed_mmS <= DL_FDR_SPD_HI)
         AND (fAccel_mmS2 >= 10.0) AND (fAccel_mmS2 <= 5000.0)
         AND (tSettle >= T#10MS) AND (tSettle <= T#500MS);
_fSpeedEff := LIMIT(DL_FDR_SPD_LO, fSpeed_mmS, DL_FDR_SPD_HI);  // 生效速度钳制 [mm/s] / Effective speed after clamping

// 段 6｜失能闸：立即停止受理，相位回空闲（不锁存故障）
IF NOT bEnable THEN
    _eState := E_DL_FeederState.eIdle;              // 相位回空闲 / Phase back to idle
    eErr := DL_FDR_READY;                           // 失能为正常停机，只回就绪码 / Disable is a normal stop, ready code only
ELSE

    // 段 7｜送料状态机（ENUM + CASE + ELSE 兜底）
    CASE _eState OF

        E_DL_FeederState.eIdle:                     // 空闲：受理请求沿 + 参数与上限校验
            IF _rtrigIndex.Q THEN
                IF NOT _bParamOk THEN
                    eErr := DL_FDR_CFG_BAD;         // 故障级：组态非法 / Fault, bad configuration
                    _uLatchCode := DL_FDR_CFG_BAD;
                    _bFaultLatch := TRUE;
                    bError := TRUE;
                    _eState := E_DL_FeederState.eFault;
                ELSE
                    _fAccumNew := fTrimAccum_mm + (fMarkOffset_mm * fTrimGain);   // 拟施加累计补偿 [mm] / Trim accumulation to be applied
                    IF (ABS(_fAccumNew) > fTrimAccumMax_mm) THEN
                        eErr := DL_FDR_ACCUM_MAX;   // 故障级：累计补偿越上限，停送 / Fault, trim accumulation beyond the limit, feeding stopped
                        _uLatchCode := DL_FDR_ACCUM_MAX;
                        _bFaultLatch := TRUE;
                        bError := TRUE;
                        _eState := E_DL_FeederState.eFault;
                    ELSE
                        _fStepRaw := fPitch_mm + (fMarkOffset_mm * fTrimGain);         // 补偿后步距 [mm] / Step distance after trim
                        _fStepEff := _fStepRaw;                                       // 生效步距初值 [mm] / Effective step initial value
                        IF _fStepRaw < (fPitch_mm * DL_FDR_STEP_LO_K) THEN
                            _fStepEff := fPitch_mm * DL_FDR_STEP_LO_K;                // 下限钳制（防倒料）[mm] / Lower clamp, prevents reverse feeding
                            eErr := DL_FDR_CLAMP;                                     // 信息级：步距已钳制 / Info, step distance clamped
                        END_IF
                        IF _fStepRaw > (fPitch_mm * DL_FDR_STEP_HI_K) THEN
                            _fStepEff := fPitch_mm * DL_FDR_STEP_HI_K;                // 上限钳制（防冲料）[mm] / Upper clamp, prevents overshoot feeding
                            eErr := DL_FDR_CLAMP;                                     // 信息级：步距已钳制 / Info, step distance clamped
                        END_IF
                        IF ABS(_fStepEff - _fStepRaw) < DL_FDR_EPS THEN
                            eErr := DL_FDR_READY;                                     // 未钳制：就绪码 / No clamping, ready code
                        END_IF
                        fStepCmd_mm := _fStepEff;                                     // 本次步距出口 [mm] / Step distance output
                        IF iAxis.MoveRelative(_fStepEff, _fSpeedEff) THEN
                            _bIssueScan := TRUE;                                      // 派单当拍不判就绪 / Readiness is not judged in the dispatch scan
                            bBusy := TRUE;
                            _eState := E_DL_FeederState.eIndexing;                    // 进入送料相 / Enter the indexing phase
                        ELSE
                            eErr := DL_FDR_AXIS_REJ;                                  // 故障级：轴拒绝指令 / Fault, the axis rejected the command
                            _uLatchCode := DL_FDR_AXIS_REJ;
                            _bFaultLatch := TRUE;
                            bError := TRUE;
                            _eState := E_DL_FeederState.eFault;
                        END_IF
                    END_IF
                END_IF
            END_IF

        E_DL_FeederState.eIndexing:                 // 送料中：请求一律丢弃（不排队），等轴就绪
            bBusy := TRUE;
            IF _bIssueScan THEN
                _bIssueScan := FALSE;                   // 派单拍已过，下一拍开始判就绪 / The dispatch scan has passed, readiness is judged from the next scan
            ELSIF iAxis.bReady THEN
                _eState := E_DL_FeederState.eSettling;  // 轴就绪：进入停稳确认 / Axis ready, enter the settle phase
            END_IF

        E_DL_FeederState.eSettling:                 // 停稳确认：计时满即完成
            bBusy := TRUE;
            IF _tonSettle.Q THEN
                uIndexCnt := uIndexCnt + 1;             // 累计送料次数 +1 [次] / Index count incremented
                bDone := TRUE;                          // 单拍完成脉冲（下一拍段 1 预清即自清） / One-scan completion pulse, self-cleared in the next scan
                eErr := DL_FDR_READY;                   // 就绪/完成码 / Ready or completion code
                bBusy := FALSE;
                _eState := E_DL_FeederState.eIdle;      // 回空闲 / Back to idle
            END_IF

        E_DL_FeederState.eFault:                    // 故障：锁存码保持，仅使能沿重启
            bBusy := FALSE;
            eErr := _uLatchCode;                        // 锁存码回放 / Replay the latch code
            bError := TRUE;                             // 故障级标志保持 / Fault flag held

        ELSE
            // 非法状态兜底（故障级，组态非法码承载）
            eErr := DL_FDR_CFG_BAD;                     // 故障级：非法相位 / Fault, illegal phase
            _uLatchCode := DL_FDR_CFG_BAD;
            _bFaultLatch := TRUE;
            bError := TRUE;
            bBusy := FALSE;
            _eState := E_DL_FeederState.eFault;

    END_CASE
END_IF

// 段 8｜累计补偿出口单点写入（全件唯一写点，禁两处赋值）
fTrimAccum_mm := _fAccumNew;                        // 累计补偿出口 [mm] / Trim accumulation output in millimetres
END_FUNCTION_BLOCK

(* ---- FB_DL_StepperXyzGantry.st ---- *)
(*==============================================================================
 * 组件名称 (Component)  : FB_DL_StepperXyzGantry
 * 所属子库 (Sublibrary) : DL_Motion
 * 当前版本 (Version)    : 1.0.1
 * 兼容性 (Platform)     : CODESYS 3.5 / TwinCAT 3 / 汇川 InoProShop（纯标准元素，零方言）
 * 功能描述 (Function)   : 三轴步进开环龙门点位运动。启动沿先做参数与软限位预检，预检
 *                         不过则一轴都不动；预检通过后按 X→Y→Z 逐轴派发相对位移，单轴
 *                         就绪即推进下一轴，每轴独立超时；三轴落定后汇总三类落点最大偏差
 *                         并给单拍完成脉冲。不做插补、不做闭环反馈、不做回零、不排队多条
 *                         目标（运行中新目标被忽略，需等待完成或中止）。
 *                         说明：接口契约 I_DL_StepperOpenLoop.MoveRelative 只接受距离与
 *                         速度，加速度由实现块组态规划，故 fAccel_mmS2 仅参与参数门禁
 *                         校验，不向下转发（规格口径已在本行登记）。
 * 溯源 (Origin)         : 道莅 clean-room 防御性实现
 * 本文件内含 (Contains) : TYPE E_DL_GantryState / FUNCTION_BLOCK FB_DL_StepperXyzGantry
 * 依赖 (Depends)        : DL_Device/I_DL_StepperOpenLoop（只调用契约方法，不复制其内核）
 * 红线自检 (Redline)    : 无外部全局变量、无硬件地址直引 ｜ 全变量中英双语同行注释
 *                         参考判空 + 参数域闸 + 软限位预检三重防御 ｜ 浮点比较用容差
 *                         非有限用自反比较 ｜ 枚举显式赋值 ｜ 超时定时器与沿检测无条件
 *                         周期刷新 ｜ CASE 含 ELSE 兜底
 * 错误码表 (Codes)      : 16#0004_0327 就绪（禁用/空闲/本拍无事件）
 *                         16#0004_0328 故障级 指令未被受理（参数域非法、轴索引越界、轴
 *                                    拒绝指令、状态机非法兜底）。反证句：轴拒绝与参数非法
 *                                    在输出侧同为「本拍无运动」，不可由 0329/032A 区分，
 *                                    故合并成一码并在头注释逐条列出四种来源
 *                         16#0004_0329 故障级 目标超软限位，启动沿前预检拒绝（一轴都不动）
 *                         16#0004_032A 故障级 单轴到位异常（超时或落点超公差），后续轴
 *                                    不再派单，当前轴受控停车
 *                         16#0004_032B 预留：本版不发码（下一轮区间起点，禁止回填）
 * 修订历史 (Revision)   : 2026-11-17  v1.0.0  首版入库 · R28 · 阶段三批 1
 *                         2026-11-17  v1.0.1  终审修复：空闲无事件相补发就绪码，消除「头注
 *                                    释声明 0327 覆盖空闲、实际输出 0」的口径不一致
 *                                    （仅输出侧，不动任何运动/判定语义）· R28 · 阶段四
 * 验收向量 (Acceptance) : 正向 X/Y 各 100 mm、Z 20 mm、50 mm/s、公差 0.01 → 逐轴推进、
 *                         偏差 ≤0.01 mm、bDone 单拍、16#0004_0327
 *                         反向 Z 目标 2500 mm（超 ±2000 软限位）→ 16#0004_0329 且三轴
 *                         位置一轴不变；速度给 0 → 16#0004_0328；单轴超时不返回就绪 →
 *                         16#0004_032A 且后续轴不再派单
 *============================================================================*)

(*-----------------------------------------------------------------------------
 * 枚举: E_DL_GantryState（归属本功能块，同文件发布，全库唯一定义）
 * 含义: 龙门点位相位，每个成员在 CASE 中有且仅有一个标签。
 *----------------------------------------------------------------------------*)
TYPE E_DL_GantryState :
(
    eIdle     := 0,    // 空闲：等待启动沿与预检 / Idle, waiting for the start edge and the pre-check
    eJogging  := 10,   // 逐轴推进：每拍只对当前轴派单与判到位 / Axis stepping, one axis dispatched per scan
    eSettling := 20,   // 落定汇总：算三类落点最大偏差 / Settling, computing the maximum deviation
    eDone     := 30,   // 完成：bDone 单拍脉冲 / Done, one-scan completion pulse
    eFault    := 99    // 故障：锁存码保持，仅复位沿退出 / Fault, the latch code is held until the reset edge
);
END_TYPE

FUNCTION_BLOCK FB_DL_StepperXyzGantry
VAR_INPUT
    bEnable      : BOOL := FALSE;         // 使能，FALSE 立即中止三轴 / Enable, FALSE aborts all three axes at once
    bStart       : BOOL := FALSE;         // 启动，上升沿启动一次（运行中被忽略） / Start, the rising edge starts one cycle and is ignored while moving
    bReset       : BOOL := FALSE;         // 复位，仅在故障态生效 / Reset, effective in the fault state only
    fTargetX_mm  : REAL := 0.0;           // X 轴目标位置 [mm]，域 ±2000 / X target position in millimetres, domain plus minus 2000
    fTargetY_mm  : REAL := 0.0;           // Y 轴目标位置 [mm]，域 ±2000 / Y target position in millimetres, domain plus minus 2000
    fTargetZ_mm  : REAL := 0.0;           // Z 轴目标位置 [mm]，域 ±2000 / Z target position in millimetres, domain plus minus 2000
    fSpeed_mmS   : REAL := 50.0;          // 运行速度 [mm/s]，域 1~500 / Run speed in millimetres per second, domain 1 to 500
    fAccel_mmS2  : REAL := 500.0;         // 加速度 [mm/s²]，域 10~5000（仅门禁校验） / Acceleration in millimetres per square second, domain 10 to 5000, gate check only
    fPosTol_mm   : REAL := 0.01;          // 落点公差 [mm]，域 0.001~1.0 / Position tolerance in millimetres, domain 0.001 to 1.0
    tAxisMax     : TIME := T#5S;          // 单轴到位超时 [ms]，域 100ms~60s / Per-axis settle timeout, domain 100 ms to 60 s
END_VAR
VAR_IN_OUT
    iAxisX       : I_DL_StepperOpenLoop;  // X 轴开环步进契约引用 [—] / X axis open-loop stepper contract reference
    iAxisY       : I_DL_StepperOpenLoop;  // Y 轴开环步进契约引用 [—] / Y axis open-loop stepper contract reference
    iAxisZ       : I_DL_StepperOpenLoop;  // Z 轴开环步进契约引用 [—] / Z axis open-loop stepper contract reference
END_VAR
VAR_OUTPUT
    fPosX_mm      : REAL;                 // X 轴实到位（指令推算）[mm] / X actual position in millimetres, open-loop derived
    fPosY_mm      : REAL;                 // Y 轴实到位（指令推算）[mm] / Y actual position in millimetres, open-loop derived
    fPosZ_mm      : REAL;                 // Z 轴实到位（指令推算）[mm] / Z actual position in millimetres, open-loop derived
    fErrMax_mm    : REAL;                 // 本次三类落点最大偏差 [mm] / Maximum deviation of the three axes in millimetres
    bDone         : BOOL;                 // 完成脉冲，单拍有效 / Completion pulse, valid for one scan
    bBusy         : BOOL;                 // 运行中 / Running
    bError        : BOOL;                 // 故障级标志，仅故障级码置位 / Fault-class flag, set on fault codes only
    eState        : E_DL_GantryState;     // 龙门相位 [—] / Gantry phase
    eErr          : UDINT;                // 错误码，段位 16#0004_xxxx / Error code in segment 16#0004_xxxx
END_VAR
VAR
    _eState       : E_DL_GantryState := E_DL_GantryState.eIdle; // 当前相位 / Current phase
    _bInit        : BOOL := FALSE;        // 首扫标志，取非判定 / First-scan flag, tested negated
    _bRefOk       : BOOL;                 // 三轴契约引用均有效标志 / All three contract references valid
    _bParamOk     : BOOL;                 // 参数门禁通过标志 / Parameter gate pass flag
    _bSoftOk      : BOOL;                 // 软限位预检通过标志 / Soft limit pre-check pass flag
    _bIssued      : BOOL;                 // 当前轴已派单标志（换轴前必清） / Current axis dispatched flag, cleared before switching axis
    _bIssueScan   : BOOL;                 // 派单当拍标志（本拍不判到位，防同拍假到位） / Dispatch scan flag, arrival is not judged in the dispatch scan
    _bSkip        : BOOL;                 // 当前轴零位移跳过标志 / Current axis skipped because the distance is zero
    _bArrived     : BOOL;                 // 当前轴就绪标志 / Current axis ready flag
    _bFaultLatch  : BOOL;                 // 故障锁存标志 / Fault latch flag
    _bAbortDone   : BOOL;                 // 失能中止已发标志（单发化） / Abort already issued flag, issued once
    _uAxisIdx     : UINT := 1;            // 当前轴索引，1=X 2=Y 3=Z / Current axis index, 1 for X, 2 for Y, 3 for Z
    _uLatchCode   : UDINT;                // 锁存码载体 / Latch code carrier
    _fAct         : REAL;                 // 当前轴回读位置 [mm] / Current axis read-back position in millimetres
    _fSpeedEff    : REAL := 50.0;         // 生效速度（下限兜底）[mm/s] / Effective speed with a lower bound guard
    _fTolEff      : REAL := 0.01;         // 生效公差（下限兜底）[mm] / Effective tolerance with a lower bound guard
    _tAxisMaxEff  : TIME := T#5S;         // 生效单轴超时（域钳制后） / Effective per-axis timeout after clamping
    _afTgt        : ARRAY[1..3] OF REAL;  // 三轴目标位置表 [mm] / Target position table of the three axes
    _afDist       : ARRAY[1..3] OF REAL;  // 三轴待走距离表 [mm] / Pending distance table of the three axes
    _afDev        : ARRAY[1..3] OF REAL;  // 三轴落点偏差表 [mm] / Deviation table of the three axes
    _rtrigStart   : R_TRIG;               // 启动上升沿 / Rising edge of the start command
    _rtrigReset   : R_TRIG;               // 复位上升沿 / Rising edge of the reset command
    _tonAxis      : TON;                  // 单轴到位超时计时 / Per-axis settle timeout timer
END_VAR
VAR CONSTANT
    DL_GTY_READY     : UDINT := 16#0004_0327;  // 就绪码 / Ready code
    DL_GTY_REJECT    : UDINT := 16#0004_0328;  // 故障级指令未受理码 / Fault code for a rejected command
    DL_GTY_LIMIT     : UDINT := 16#0004_0329;  // 故障级超软限位码 / Fault code for a soft limit violation
    DL_GTY_AXIS_BAD  : UDINT := 16#0004_032A;  // 故障级单轴到位异常码 / Fault code for an abnormal axis settle
    DL_GTY_SOFT_MM   : REAL := 2000.0;         // 软限位绝对值 [mm] / Absolute soft limit in millimetres
    DL_GTY_EPS_MM    : REAL := 0.001;          // 零位移判定容差 [mm] / Zero-distance tolerance in millimetres
    DL_GTY_SPD_LO    : REAL := 1.0;            // 速度下限 [mm/s] / Speed lower bound
    DL_GTY_SPD_HI    : REAL := 500.0;          // 速度上限 [mm/s] / Speed upper bound
    DL_GTY_ACC_LO    : REAL := 10.0;           // 加速度下限 [mm/s²] / Acceleration lower bound
    DL_GTY_ACC_HI    : REAL := 5000.0;         // 加速度上限 [mm/s²] / Acceleration upper bound
    DL_GTY_TOL_LO    : REAL := 0.001;          // 公差下限 [mm] / Tolerance lower bound
    DL_GTY_TOL_HI    : REAL := 1.0;            // 公差上限 [mm] / Tolerance upper bound
END_VAR

// 段 1｜输出与单拍标志预置（每拍重算，禁跨拍残留）
bDone := FALSE;                                     // 完成脉冲预清 / Completion pulse pre-cleared
bBusy := FALSE;                                     // 运行标志预清 / Busy flag pre-cleared
bError := FALSE;                                    // 故障标志预清 / Fault flag pre-cleared
eErr := 0;                                          // 错误码预清 / Error code pre-cleared
_bIssueScan := FALSE;                               // 派单当拍标志预清 / Dispatch scan flag pre-cleared
_bArrived := FALSE;                                 // 到位标志预清 / Arrival flag pre-cleared
_fAct := 0.0;                                       // 回读位置预清 / Read-back position pre-cleared

// 段 2｜沿检测无条件周期刷新（严禁置于分支内）
_rtrigStart(CLK := bStart);                         // 启动沿 / Start edge
_rtrigReset(CLK := bReset);                         // 复位沿 / Reset edge

// 段 3｜超时定时器无条件周期刷新（仅推进态且已派单时计时）
_tonAxis(IN := (_eState = E_DL_GantryState.eJogging) AND _bIssued, PT := _tAxisMaxEff);

// 段 4｜首扫初始化（判据取非，R19）
IF NOT _bInit THEN
    _eState := E_DL_GantryState.eIdle;              // 相位待机起步 / Phase starts idle
    _uAxisIdx := 1;                                 // 轴索引起步为 X / Axis index starts at X
    _bInit := TRUE;                                 // 首扫只做一次 / The first scan runs once
END_IF

// 段 5｜契约引用有效性（任一未注入即拒绝启动，不产生误动作）
_bRefOk := NOT ((iAxisX = 0) OR (iAxisY = 0) OR (iAxisZ = 0));

// 段 6｜参数门禁逐拍重算（非有限用自反比较，禁近似阈值）
_bParamOk := _bRefOk
         AND NOT ((fSpeed_mmS <> fSpeed_mmS) OR ((fSpeed_mmS - fSpeed_mmS) <> (fSpeed_mmS - fSpeed_mmS)))
         AND NOT ((fAccel_mmS2 <> fAccel_mmS2) OR ((fAccel_mmS2 - fAccel_mmS2) <> (fAccel_mmS2 - fAccel_mmS2)))
         AND NOT ((fPosTol_mm <> fPosTol_mm) OR ((fPosTol_mm - fPosTol_mm) <> (fPosTol_mm - fPosTol_mm)))
         AND (fSpeed_mmS >= DL_GTY_SPD_LO) AND (fSpeed_mmS <= DL_GTY_SPD_HI)
         AND (fAccel_mmS2 >= DL_GTY_ACC_LO) AND (fAccel_mmS2 <= DL_GTY_ACC_HI)
         AND (fPosTol_mm >= DL_GTY_TOL_LO) AND (fPosTol_mm <= DL_GTY_TOL_HI)
         AND (tAxisMax >= T#100MS) AND (tAxisMax <= T#60S);
_fSpeedEff := LIMIT(DL_GTY_SPD_LO, fSpeed_mmS, DL_GTY_SPD_HI);   // 生效速度钳制 [mm/s] / Effective speed after clamping
_fTolEff := LIMIT(DL_GTY_TOL_LO, fPosTol_mm, DL_GTY_TOL_HI);     // 生效公差钳制 [mm] / Effective tolerance after clamping
_tAxisMaxEff := LIMIT(T#100MS, tAxisMax, T#60S);                  // 生效超时钳制 [ms] / Effective timeout after clamping

// 段 7｜目标与软限位预检（超限位则启动沿前一拍即拒绝，一轴不动）
_afTgt[1] := fTargetX_mm;                           // X 目标入表 [mm] / X target into the table
_afTgt[2] := fTargetY_mm;                           // Y 目标入表 [mm] / Y target into the table
_afTgt[3] := fTargetZ_mm;                           // Z 目标入表 [mm] / Z target into the table
_bSoftOk := TRUE;                                   // 软限位预检假设成立 / Assume the soft limit pre-check passes
IF (fTargetX_mm <> fTargetX_mm) OR ((fTargetX_mm - fTargetX_mm) <> (fTargetX_mm - fTargetX_mm)) THEN
    _bSoftOk := FALSE;                              // X 目标非有限 / X target not finite
END_IF
IF (fTargetY_mm <> fTargetY_mm) OR ((fTargetY_mm - fTargetY_mm) <> (fTargetY_mm - fTargetY_mm)) THEN
    _bSoftOk := FALSE;                              // Y 目标非有限 / Y target not finite
END_IF
IF (fTargetZ_mm <> fTargetZ_mm) OR ((fTargetZ_mm - fTargetZ_mm) <> (fTargetZ_mm - fTargetZ_mm)) THEN
    _bSoftOk := FALSE;                              // Z 目标非有限 / Z target not finite
END_IF
IF (ABS(fTargetX_mm) > DL_GTY_SOFT_MM) THEN
    _bSoftOk := FALSE;                              // X 超软限位 / X beyond the soft limit
END_IF
IF (ABS(fTargetY_mm) > DL_GTY_SOFT_MM) THEN
    _bSoftOk := FALSE;                              // Y 超软限位 / Y beyond the soft limit
END_IF
IF (ABS(fTargetZ_mm) > DL_GTY_SOFT_MM) THEN
    _bSoftOk := FALSE;                              // Z 超软限位 / Z beyond the soft limit
END_IF

// 段 8｜实际位置回读（引用有效时每拍刷新，禁用时保持上次值）
IF _bRefOk THEN
    fPosX_mm := iAxisX.fPosition;                   // X 实到位 [mm] / X actual position
    fPosY_mm := iAxisY.fPosition;                   // Y 实到位 [mm] / Y actual position
    fPosZ_mm := iAxisZ.fPosition;                   // Z 实到位 [mm] / Z actual position
ELSE
    fPosX_mm := 0.0;                                // 引用无效：输出置 0 并随故障码上报 / Invalid reference, outputs zeroed and reported with the fault code
    fPosY_mm := 0.0;
    fPosZ_mm := 0.0;
    _bSoftOk := FALSE;                              // 引用无效一并拒绝启动 / An invalid reference also blocks the start
END_IF

// 段 9｜失能立即中止（单发停车，不清位置；状态回空闲）
IF NOT bEnable THEN
    IF NOT _bAbortDone THEN
        _bAbortDone := TRUE;                        // 中止只发一次 / The abort is issued once
        IF _bRefOk THEN
            iAxisX.Stop();                          // X 受控停车 / X controlled stop
            iAxisY.Stop();                          // Y 受控停车 / Y controlled stop
            iAxisZ.Stop();                          // Z 受控停车 / Z controlled stop
        END_IF
    END_IF
    _bIssued := FALSE;                              // 派单标志清 / Dispatch flag cleared
    _uAxisIdx := 1;                                 // 轴索引回 X / Axis index back to X
    _eState := E_DL_GantryState.eIdle;              // 相位回空闲 / Phase back to idle
    eErr := DL_GTY_READY;                           // 失能为正常停机，只回就绪码 / Disable is a normal stop, ready code only
ELSE
    _bAbortDone := FALSE;                           // 使能期清中止标志 / Abort flag cleared while enabled
END_IF

// 段 10｜龙门点位状态机（ENUM + CASE + ELSE 兜底）
CASE _eState OF

    E_DL_GantryState.eIdle:                         // 空闲：等启动沿 + 三重预检
        IF _rtrigStart.Q AND bEnable THEN
            _bFaultLatch := FALSE;                  // 新启动沿为锁存解除路径 / A new start edge is the latch release path
            _uLatchCode := 0;                       // 锁存码清 / Latch code cleared
            _bIssued := FALSE;                      // 派单标志清 / Dispatch flag cleared
            _uAxisIdx := 1;                         // 从 X 轴起步 / Start from the X axis
            _afDev[1] := 0.0;                       // 偏差表清零 [mm] / Deviation table cleared
            _afDev[2] := 0.0;
            _afDev[3] := 0.0;
            fErrMax_mm := 0.0;                      // 本次最大偏差清 [mm] / Maximum deviation cleared
            IF NOT _bRefOk THEN
                eErr := DL_GTY_REJECT;              // 故障级：契约引用未注入 / Fault, a contract reference is missing
                _uLatchCode := DL_GTY_REJECT;
                _bFaultLatch := TRUE;
                bError := TRUE;
                _eState := E_DL_GantryState.eFault;
            ELSIF NOT _bParamOk THEN
                eErr := DL_GTY_REJECT;              // 故障级：参数域非法 / Fault, parameters out of domain
                _uLatchCode := DL_GTY_REJECT;
                _bFaultLatch := TRUE;
                bError := TRUE;
                _eState := E_DL_GantryState.eFault;
            ELSIF NOT _bSoftOk THEN
                eErr := DL_GTY_LIMIT;               // 故障级：超软限位，一轴都不动 / Fault, beyond the soft limit, no axis moves
                _uLatchCode := DL_GTY_LIMIT;
                _bFaultLatch := TRUE;
                bError := TRUE;
                _eState := E_DL_GantryState.eFault;
            ELSE
                _afDist[1] := _afTgt[1] - iAxisX.fPosition;   // X 待走距离 [mm] / X pending distance
                _afDist[2] := _afTgt[2] - iAxisY.fPosition;   // Y 待走距离 [mm] / Y pending distance
                _afDist[3] := _afTgt[3] - iAxisZ.fPosition;   // Z 待走距离 [mm] / Z pending distance
                IF (ABS(_afDist[1]) <= DL_GTY_EPS_MM) AND (ABS(_afDist[2]) <= DL_GTY_EPS_MM) AND (ABS(_afDist[3]) <= DL_GTY_EPS_MM) THEN
                    _eState := E_DL_GantryState.eDone;        // 三轴零位移直通完成（零位移指令在部分平台挂死） / All distances zero, finish directly
                ELSE
                    _eState := E_DL_GantryState.eJogging;     // 进入逐轴推进 / Enter the per-axis stepping phase
                END_IF
            END_IF
        ELSE
            eErr := DL_GTY_READY;                       // 空闲无事件：回就绪码（对齐码表口径） / Idle without an event, ready code
        END_IF

    E_DL_GantryState.eJogging:                      // 逐轴推进：派单一次，判就绪或超时
        bBusy := TRUE;
        IF (_uAxisIdx < 1) OR (_uAxisIdx > 3) THEN
            eErr := DL_GTY_REJECT;                  // 故障级：轴索引越界 / Fault, axis index out of range
            _uLatchCode := DL_GTY_REJECT;
            _bFaultLatch := TRUE;
            bError := TRUE;
            bBusy := FALSE;
            _eState := E_DL_GantryState.eFault;
        ELSE
            // 派单（每轴只发一次；零位移轴跳过，不派单）
            IF NOT _bIssued THEN
                _bSkip := FALSE;                    // 跳过标志预清 / Skip flag pre-cleared
                CASE _uAxisIdx OF
                    1:
                        IF ABS(_afDist[1]) <= DL_GTY_EPS_MM THEN
                            _bSkip := TRUE;         // X 零位移跳过 / X skipped, zero distance
                        ELSE
                            _bIssued := iAxisX.MoveRelative(_afDist[1], _fSpeedEff);  // X 相对位移派发 / X relative move dispatched
                            _bIssueScan := TRUE;    // 派单当拍不判到位 / Arrival is not judged in the dispatch scan
                        END_IF
                    2:
                        IF ABS(_afDist[2]) <= DL_GTY_EPS_MM THEN
                            _bSkip := TRUE;         // Y 零位移跳过 / Y skipped, zero distance
                        ELSE
                            _bIssued := iAxisY.MoveRelative(_afDist[2], _fSpeedEff);  // Y 相对位移派发 / Y relative move dispatched
                            _bIssueScan := TRUE;    // 派单当拍不判到位 / Arrival is not judged in the dispatch scan
                        END_IF
                    3:
                        IF ABS(_afDist[3]) <= DL_GTY_EPS_MM THEN
                            _bSkip := TRUE;         // Z 零位移跳过 / Z skipped, zero distance
                        ELSE
                            _bIssued := iAxisZ.MoveRelative(_afDist[3], _fSpeedEff);  // Z 相对位移派发 / Z relative move dispatched
                            _bIssueScan := TRUE;    // 派单当拍不判到位 / Arrival is not judged in the dispatch scan
                        END_IF
                    ELSE
                        _bSkip := FALSE;            // 非 1~3 索引：交由上层索引防御拦截 / Other indices are rejected by the range guard above
                END_CASE
                IF (NOT _bIssued) AND (NOT _bSkip) THEN
                    eErr := DL_GTY_REJECT;          // 故障级：轴拒绝指令 / Fault, the axis rejected the command
                    _uLatchCode := DL_GTY_REJECT;
                    _bFaultLatch := TRUE;
                    bError := TRUE;
                    bBusy := FALSE;
                    _eState := E_DL_GantryState.eFault;
                ELSIF _bSkip THEN
                    _uAxisIdx := _uAxisIdx + 1;     // 零位移轴直接推进 / Advance past the zero-distance axis
                    IF _uAxisIdx > 3 THEN
                        _eState := E_DL_GantryState.eSettling;   // 三轴已处理完 / All three axes handled
                    END_IF
                END_IF
            END_IF

            // 到位判定（派单当拍跳过，防同拍假到位）
            IF (_eState = E_DL_GantryState.eJogging) AND _bIssued AND (NOT _bIssueScan) THEN
                CASE _uAxisIdx OF
                    1:
                        _bArrived := iAxisX.bReady;         // X 就绪（空闲且无故障） / X ready, idle and fault free
                        _fAct := iAxisX.fPosition;          // X 回读位置 [mm] / X read-back position
                    2:
                        _bArrived := iAxisY.bReady;         // Y 就绪 / Y ready
                        _fAct := iAxisY.fPosition;          // Y 回读位置 [mm] / Y read-back position
                    3:
                        _bArrived := iAxisZ.bReady;         // Z 就绪 / Z ready
                        _fAct := iAxisZ.fPosition;          // Z 回读位置 [mm] / Z read-back position
                    ELSE
                        _bArrived := FALSE;                 // 非法索引不判到位 / No arrival judgement on an illegal index
                        _fAct := 0.0;
                END_CASE
                _afDev[_uAxisIdx] := ABS(_afTgt[_uAxisIdx] - _fAct);   // 当前轴落点偏差 [mm] / Deviation of the current axis
                IF _tonAxis.Q THEN
                    _bIssued := FALSE;                  // 超时：清派单，不再发新指令 / Timeout, clear the dispatch and issue nothing further
                    CASE _uAxisIdx OF
                        1: iAxisX.Stop();               // X 受控停车 / X controlled stop
                        2: iAxisY.Stop();               // Y 受控停车 / Y controlled stop
                        3: iAxisZ.Stop();               // Z 受控停车 / Z controlled stop
                        ELSE _bArrived := FALSE;        // 非法索引无停车对象 / No stop target for an illegal index
                    END_CASE
                    eErr := DL_GTY_AXIS_BAD;            // 故障级：单轴到位超时 / Fault, per-axis settle timeout
                    _uLatchCode := DL_GTY_AXIS_BAD;
                    _bFaultLatch := TRUE;
                    bError := TRUE;
                    bBusy := FALSE;
                    _eState := E_DL_GantryState.eFault;
                ELSIF _bArrived THEN
                    IF _afDev[_uAxisIdx] > _fTolEff THEN
                        eErr := DL_GTY_AXIS_BAD;        // 故障级：落点超公差（与超时同族） / Fault, position deviation beyond tolerance
                        _uLatchCode := DL_GTY_AXIS_BAD;
                        _bFaultLatch := TRUE;
                        bError := TRUE;
                        bBusy := FALSE;
                        _eState := E_DL_GantryState.eFault;
                    ELSE
                        _bIssued := FALSE;              // 换轴前清上一轴派单标志（R27 跨轴标志） / Clear the dispatch flag before switching axis
                        _uAxisIdx := _uAxisIdx + 1;     // 推进下一轴 / Advance to the next axis
                        IF _uAxisIdx > 3 THEN
                            _eState := E_DL_GantryState.eSettling;   // 三轴落定 / All three axes settled
                        END_IF
                    END_IF
                END_IF
            END_IF
        END_IF

    E_DL_GantryState.eSettling:                     // 落定汇总：三类落点最大偏差
        bBusy := TRUE;
        IF _bRefOk THEN
            _afDev[1] := ABS(_afTgt[1] - iAxisX.fPosition);   // X 落点偏差 [mm] / X deviation
            _afDev[2] := ABS(_afTgt[2] - iAxisY.fPosition);   // Y 落点偏差 [mm] / Y deviation
            _afDev[3] := ABS(_afTgt[3] - iAxisZ.fPosition);   // Z 落点偏差 [mm] / Z deviation
        END_IF
        fErrMax_mm := _afDev[1];                    // 最大偏差初值取 X [mm] / Maximum deviation initialised with X
        IF _afDev[2] > fErrMax_mm THEN
            fErrMax_mm := _afDev[2];                // Y 更大则替换 [mm] / Replaced when Y is larger
        END_IF
        IF _afDev[3] > fErrMax_mm THEN
            fErrMax_mm := _afDev[3];                // Z 更大则替换 [mm] / Replaced when Z is larger
        END_IF
        _eState := E_DL_GantryState.eDone;          // 下一拍进入完成相 / Enter the done phase on the next scan

    E_DL_GantryState.eDone:                         // 拍 N 进入：三轴到位；本拍行为：置 bDone 单拍脉冲；
        bDone := TRUE;                              // 拍 N+1 转出并回空闲，段 1 预清即自清（R24 三律） / The pulse self-clears in the next scan
        bBusy := FALSE;
        eErr := DL_GTY_READY;                       // 正常完成只回就绪码 / A normal completion reports the ready code only
        _eState := E_DL_GantryState.eIdle;          // 相位回空闲 / Phase back to idle

    E_DL_GantryState.eFault:                        // 故障：锁存码保持，仅复位沿退出
        bBusy := FALSE;
        eErr := _uLatchCode;                        // 锁存码回放 / Replay the latch code
        bError := TRUE;                             // 故障级标志保持 / Fault flag held
        IF _rtrigReset.Q THEN
            IF _bRefOk THEN
                iAxisX.Reset();                     // X 故障复位 / X fault reset
                iAxisY.Reset();                     // Y 故障复位 / Y fault reset
                iAxisZ.Reset();                     // Z 故障复位 / Z fault reset
            END_IF
            _bFaultLatch := FALSE;                  // 锁存解除 / Latch released
            _uLatchCode := 0;                       // 锁存码清 / Latch code cleared
            _bIssued := FALSE;                      // 派单标志清 / Dispatch flag cleared
            _uAxisIdx := 1;                         // 轴索引回 X / Axis index back to X
            eErr := DL_GTY_READY;                   // 复位后回就绪码 / Ready code after the reset
            bError := FALSE;
            _eState := E_DL_GantryState.eIdle;      // 回空闲需新启动沿 / Back to idle, a new start edge is required
        END_IF

    ELSE
        // 非法状态兜底（故障级，指令未受理码承载）
        eErr := DL_GTY_REJECT;                      // 故障级：非法相位 / Fault, illegal phase
        _uLatchCode := DL_GTY_REJECT;
        _bFaultLatch := TRUE;
        bError := TRUE;
        bBusy := FALSE;
        _bIssued := FALSE;
        _eState := E_DL_GantryState.eFault;

END_CASE

eState := _eState;                                  // 相位出口镜像（只读引脚） / Phase mirrored to the output pin
END_FUNCTION_BLOCK

(* ---- FB_DL_StepperZLiftMicron.st ---- *)
(*==============================================================================
 * 组件名称 (Component)  : FB_DL_StepperZLiftMicron
 * 所属子库 (Sublibrary) : DL_Motion
 * 当前版本 (Version)    : 1.0.0
 * 兼容性 (Platform)     : CODESYS 3.5 / TwinCAT 3 / 汇川 InoProShop / Machine Expert
 *                         仅依赖纯 IEC 61131-3 标准元素，零厂商方言
 * 功能描述 (Function)   : Z 轴微米级步进升降：细分当量组态（um/步）+ 相对目标
 *                         微动 + 软限位行程拦截。目标先 ROUND 换算步数（防浮点
 *                         累积）并做步数溢出检测（> 1e7 拒绝）；软限位预检先行；
 *                         运动中越限立即急停拦截；步脉冲经 TP 成形，位置以
 *                         LREAL 累加防微米级累积误差。
 * 溯源 (Origin)         : 道莅 clean-room 防御性实现
 * 本文件内含 (Contains) : TYPE E_DL_StepZState / TYPE E_DL_StepZErr /
 *                         FUNCTION_BLOCK FB_DL_StepperZLiftMicron
 * 依赖 (Depends)        : DL_MathData/FC_DL_DintMsToTime、DL_MathData/FC_DL_TimeToLrealSec
 * 红线自检 (Redline)    : 无外部全局变量、无硬件地址直引 ｜ 全变量中英双语同行注释
 *                         当量下限防除零 + 步数溢出检测 + 速度钳位 + 非有限防御 ｜
 *                         枚举成员全部显式赋值 ｜ TP/TON/R_TRIG 每周期无条件调用 ｜
 *                         状态机 CASE 含 ELSE 兜底 ｜ 位置累加用 LREAL
 * 错误码表 (Codes)      : 16#0004_0322 就绪
 *                         16#0004_0323 故障级 配置非法（当量/速度/限位组态，共用反证句）
 *                         16#0004_0324 故障级 目标超软限位或步数溢出（拒绝启动，共用反证句）
 *                         16#0004_0325 故障级 运动中限位拦截(急停)
 *                         16#0004_0326 到位
 * 修订历史 (Revision)   : 2026-11-17  v1.0.0  首版入库 · R27 · 阶段三批 3
 * 验收向量 (Acceptance) : 当量 0.5 um/步，目标 +100 um → 200 步；到位 0326；
 *                         目标超上限 → 0324 拒绝；运动中 fPosNow 越限 → 0325 急停
 *============================================================================*)

(*-----------------------------------------------------------------------------
 * 枚举: E_DL_StepZState（归属 DL_Motion，步进状态机状态）
 *----------------------------------------------------------------------------*)
TYPE E_DL_StepZState :
(
    eIdle    := 0,    // 就绪待启动 / Idle, waiting for a start
    eMoving  := 10,   // 步进运动中（TP 成形步脉冲）/ Stepping, TP-formed pulses
    eDone    := 20,   // 到位（保持至下一次启动）/ In position, held until next start
    eFault   := 99    // 故障兜底态（急停后保持）/ Fault fallback, held after e-stop
);
END_TYPE

(*-----------------------------------------------------------------------------
 * 枚举: E_DL_StepZErr（归属 DL_Motion，与 FB_DL_StepperZLiftMicron 同文件）
 *----------------------------------------------------------------------------*)
TYPE E_DL_StepZErr :
(
    eReady     := 16#0004_0322,   // 就绪 / Ready
    eConfigBad := 16#0004_0323,   // 故障级：配置非法（当量/速度/限位组态）/ Fault: illegal configuration
    eTargetBad := 16#0004_0324,   // 故障级：目标超软限位或步数溢出 / Fault: target beyond soft limit or step overflow
    eLimitHit  := 16#0004_0325,   // 故障级：运动中限位拦截（急停）/ Fault: limit hit in motion, e-stop
    eInPos     := 16#0004_0326    // 到位 / In position
);
END_TYPE

(*==============================================================================
 * 功能块: FB_DL_StepperZLiftMicron
 * 调用约定: 每个扫描周期无条件调用一次；tSampleTime 注入真实任务间隔。
 *============================================================================*)
FUNCTION_BLOCK FB_DL_StepperZLiftMicron
VAR_INPUT
    fUmPerStep  : REAL;                // 细分当量 [微米每步]，有效域 0.01~100 / Micrometers per step, subdivision config
    fTargetUm   : REAL;                // 目标位置 [微米]（绝对目标）/ Target position [um]
    fUpLimit_um : REAL;                // 软限位上限 [微米] / Soft limit upper [um]
    fLoLimit_um : REAL;                // 软限位下限 [微米] / Soft limit lower [um]
    fSpeedPps   : UDINT;               // 速度 [步每秒]，有效域 1~100000 / Speed [steps per second]
    bStartMove  : BOOL;                // 启动微动（上升沿）/ Start move trigger, rising edge
    bReset      : BOOL;                // 故障复位（上升沿）/ Fault reset, rising edge
    tSampleTime : TIME := T#1MS;       // 采样周期，调用方注入 / Sample period, caller-injected
END_VAR
VAR_OUTPUT
    fPosNow_um  : LREAL;               // 当前位置 [微米]（LREAL 累加防累积误差）/ Current position [um], LREAL accumulation
    bMoving     : BOOL;                // 运动中标志 / Moving flag
    bStepPulse  : BOOL;                // 步脉冲输出（TP 成形）/ Step pulse output, TP-formed
    bLimitHit   : BOOL;                // 限位拦截标志（锁存至复位）/ Limit-hit flag, latched until reset
    eErr        : E_DL_StepZErr;       // 错误码 / Error code
    eState      : E_DL_StepZState;     // 步进状态机当前状态 / Stepper state
END_VAR
VAR
    fbStartTrig : R_TRIG;              // 启动沿实例（无条件调用）/ Start edge instance
    fbResetTrig : R_TRIG;              // 复位沿实例（无条件调用）/ Reset edge instance
    fbPulse     : TP;                  // 步脉冲成形实例（无条件调用）/ Step pulse forming instance
    nStepsTotal : DINT;                // 本程总步数 [步]（ROUND 换算）/ Total steps this move [steps]
    nStepsDone  : DINT;                // 已发步数 [步] / Steps issued [steps]
    fStepAcc    : LREAL;               // 步数小数累积器 [步] / Fractional step accumulator [steps]
    fEquivUse   : REAL;                // 生效当量（钳位后）[微米每步] / Effective equivalence [um per step]
    fSpeedUse   : UDINT;               // 生效速度（钳位后）[步每秒] / Effective speed [steps per second]
    fUpUse      : REAL;                // 生效软限位上限 [微米] / Effective upper soft limit [um]
    fLoUse      : REAL;                // 生效软限位下限 [微米] / Effective lower soft limit [um]
    fTargetUse  : REAL;                // 生效目标（NaN 拒绝）[微米] / Effective target [um]
    fStepPulseW : TIME;                // 步脉冲宽度 [毫秒]（半步周期，委托换算）/ Step pulse width [ms] via delegate
    fDirSign    : LREAL;               // 运动方向符号（+1 上行 / -1 下行）/ Direction sign, plus up minus down
    fDtSec      : LREAL;               // 采样周期秒值（委托换算）[秒] / Sample period seconds via delegate
    bNonFin     : BOOL;                // 非有限输入汇总标志 / Non-finite input aggregate flag
    bStepReq    : BOOL;                // 步脉冲请求锁存（TP 输入源，脉宽完成后解锁）/ Step pulse request latch, released after the pulse
    uTmErr      : UDINT;               // 委托时间换算错误码（0 = 无错）/ Delegate time error id
END_VAR
VAR CONSTANT
    DL_STZ_EQUIV_MIN  : REAL := 0.01;     // 当量下限 [微米每步] / Equivalence lower bound [um per step]
    DL_STZ_EQUIV_MAX  : REAL := 100.0;    // 当量上限 [微米每步] / Equivalence upper bound [um per step]
    DL_STZ_SPEED_MIN  : UDINT := 1;       // 速度下限 [步每秒] / Speed lower bound [steps per s]
    DL_STZ_SPEED_MAX  : UDINT := 100000;  // 速度上限 [步每秒] / Speed upper bound [steps per s]
    DL_STZ_STEPS_MAX  : DINT := 10000000; // 步数溢出上限 [步] / Step overflow bound [steps]
    DL_STZ_INF_MAX    : REAL := 1.0E30;   // 非有限值判定幅值上限 / Magnitude bound for finite-value check
    DL_STZ_ZERO       : REAL := 0.0;      // 零值常量，避免裸字面量 / Zero constant
    DL_STZ_TOL        : REAL := 1.0E-6;   // 浮点比较容差 / Float comparison tolerance
END_VAR

(*------------------------------------------------------------------------------
 * 段 1｜沿检测/TP 实例每周期无条件调用（仅输入条件化）
 *----------------------------------------------------------------------------*)
fbStartTrig(CLK := bStartMove);                       // 启动沿检测无条件刷新 / start edge refreshed unconditionally
fbResetTrig(CLK := bReset);                           // 复位沿检测无条件刷新 / reset edge refreshed unconditionally
fbPulse(IN := bStepReq, PT := fStepPulseW);   // 步脉冲成形（请求锁存源，宽度为半步周期）/ step pulse formed

(*------------------------------------------------------------------------------
 * 段 2｜复位沿：故障清除回就绪（限位标志解锁）
 *----------------------------------------------------------------------------*)
IF fbResetTrig.Q THEN
    eState := E_DL_StepZState.eIdle;                 // 回就绪态 / back to idle
    eErr := E_DL_StepZErr.eReady;                    // 回就绪码 / back to ready
    bLimitHit := FALSE;                              // 限位标志解锁 / limit flag released
    bMoving := FALSE;                                // 运动标志撤 / moving dropped
END_IF

(*------------------------------------------------------------------------------
 * 段 3｜非有限值闸与配置钳位：当量/速度/限位非法 → 0323（共用反证句）
 *----------------------------------------------------------------------------*)
bNonFin := (fUmPerStep <> fUmPerStep) OR (ABS(fUmPerStep) > DL_STZ_INF_MAX)
        OR (fTargetUm  <> fTargetUm)  OR (ABS(fTargetUm)  > DL_STZ_INF_MAX)
        OR (fUpLimit_um <> fUpLimit_um) OR (ABS(fUpLimit_um) > DL_STZ_INF_MAX)
        OR (fLoLimit_um <> fLoLimit_um) OR (ABS(fLoLimit_um) > DL_STZ_INF_MAX);
IF bNonFin THEN
    eState := E_DL_StepZState.eFault;                // 进故障态 / enter fault
    eErr := E_DL_StepZErr.eConfigBad;                // 故障级：配置非法（非有限并入配置段）/ fault: config band
    bMoving := FALSE;                                // 运动撤 / moving dropped
    bStepPulse := FALSE;                             // 脉冲撤 / pulse dropped
    RETURN;
END_IF
fEquivUse := fUmPerStep;                              // 当量工作副本 / equivalence working copy
IF (fEquivUse < DL_STZ_EQUIV_MIN) OR (fEquivUse > DL_STZ_EQUIV_MAX) THEN
    eErr := E_DL_StepZErr.eConfigBad;                // 故障级：当量非法 / fault: illegal equivalence
    IF eState = E_DL_StepZState.eMoving THEN
        eState := E_DL_StepZState.eFault;            // 运动中配置突变：急停进故障态 / config change in motion: e-stop
        bMoving := FALSE;                            // 运动撤 / moving dropped
    END_IF
END_IF
fSpeedUse := fSpeedPps;                               // 速度工作副本 / speed working copy
IF (fSpeedUse < DL_STZ_SPEED_MIN) OR (fSpeedUse > DL_STZ_SPEED_MAX) THEN
    IF fSpeedUse < DL_STZ_SPEED_MIN THEN
        fSpeedUse := DL_STZ_SPEED_MIN;               // 速度下限钳位 / speed floored
    ELSE
        fSpeedUse := DL_STZ_SPEED_MAX;               // 速度上限钳位 / speed capped
    END_IF
END_IF
fUpUse := fUpLimit_um;                                // 上限工作副本 / upper working copy
fLoUse := fLoLimit_um;                                // 下限工作副本 / lower working copy
IF fLoUse >= fUpUse THEN
    eErr := E_DL_StepZErr.eConfigBad;                 // 故障级：限位组态非法（下限 >= 上限）/ fault: illegal limit config
    IF eState = E_DL_StepZState.eMoving THEN
        eState := E_DL_StepZState.eFault;            // 运动中组态突变：急停 / config change in motion: e-stop
        bMoving := FALSE;                            // 运动撤 / moving dropped
    END_IF
END_IF

(*------------------------------------------------------------------------------
 * 段 4｜速度换算：步周期 [毫秒] 与采样周期秒值（委托，防除零）
 *----------------------------------------------------------------------------*)
fStepPulseW := FC_DL_DintMsToTime(nMs := REAL_TO_DINT(500.0 / UDINT_TO_REAL(fSpeedUse)), eErr => uTmErr);   // 脉宽 = 半步周期（500/speed ms，委托换算；速度已钳位为正，除子非零）/ pulse width via delegate
IF uTmErr <> 0 THEN
    fStepPulseW := T#1MS;                             // 换算失败按 1 ms 兜底 / conversion failure falls back to 1 ms
END_IF
fDtSec := FC_DL_TimeToLrealSec(tIn := tSampleTime);   // 采样周期秒值（委托换算）/ sample period seconds via delegate
IF (fDtSec <> fDtSec) OR (fDtSec < LREAL#1.0E-6) THEN
    fDtSec := LREAL#0.001;                            // 非法采样周期按 1 ms 兜底（防除零）/ illegal sample period falls back
END_IF

(*------------------------------------------------------------------------------
 * 段 5｜启动沿：软限位预检先行 + ROUND 换算步数 + 溢出检测 → 0324 拒绝
 *----------------------------------------------------------------------------*)
IF fbStartTrig.Q AND (eState <> E_DL_StepZState.eFault) AND (eErr <> E_DL_StepZErr.eConfigBad) THEN
    fTargetUse := fTargetUm;                          // 目标工作副本 / target working copy
    IF (fTargetUse > fUpUse + DL_STZ_TOL) OR (fTargetUse < fLoUse - DL_STZ_TOL) THEN
        eErr := E_DL_StepZErr.eTargetBad;             // 故障级：目标超软限位（预检拒绝）/ fault: target beyond soft limit
    ELSE
        nStepsTotal := REAL_TO_DINT(ROUND((fTargetUse - fPosNow_um) / fEquivUse));   // ROUND 换算步数（防浮点累积）/ steps by ROUND
        IF (nStepsTotal > DL_STZ_STEPS_MAX) OR (nStepsTotal < -DL_STZ_STEPS_MAX) THEN
            eErr := E_DL_StepZErr.eTargetBad;         // 故障级：步数溢出（与超限共用 0324，反证句：同为拒绝启动+脉冲撤）/ fault: step overflow
            nStepsTotal := 0;                         // 步数清零 / steps cleared
        ELSE
            nStepsDone := 0;                          // 已发步数清零 / issued steps cleared
            fStepAcc := LREAL#0.0;                    // 小数累积器清零 / fractional accumulator cleared
            IF (fTargetUse - fPosNow_um) >= DL_STZ_ZERO THEN
                fDirSign := LREAL#1.0;                // 上行方向 / upward direction
            ELSE
                fDirSign := LREAL#-1.0;               // 下行方向 / downward direction
            END_IF
            IF nStepsTotal = 0 THEN
                eErr := E_DL_StepZErr.eInPos;         // 零步数：已在目标位 / zero steps: already in position
                eState := E_DL_StepZState.eDone;      // 进到位相 / enter done phase
            ELSE
                eState := E_DL_StepZState.eMoving;    // 启动运动 / start moving
            END_IF
        END_IF
    END_IF
END_IF

(*------------------------------------------------------------------------------
 * 段 6｜步进运动：按速度累积步数（LREAL），整数步经 TP 成形脉冲发出
 *----------------------------------------------------------------------------*)
bMoving := (eState = E_DL_StepZState.eMoving);        // 运动标志随状态 / moving follows state
bStepPulse := fbPulse.Q;                              // 脉冲输出由 TP 成形结果驱动 / pulse output driven by the TP result
IF fbPulse.Q THEN
    bStepReq := FALSE;                                // 脉宽完成：请求解锁 / pulse done: request released
END_IF
IF eState = E_DL_StepZState.eMoving THEN
    fStepAcc := fStepAcc + UDINT_TO_LREAL(fSpeedUse) * fDtSec;   // 步数累积 [步] / step accumulation
    WHILE (fStepAcc >= LREAL#1.0) AND (nStepsDone < nStepsTotal) DO
        fStepAcc := fStepAcc - LREAL#1.0;             // 消耗一个整数步 / consume one integer step
        nStepsDone := nStepsDone + 1;                 // 已发步数递增 [步] / issued steps incremented
        bStepReq := TRUE;                             // 步脉冲请求锁存（下拍 TP 成形）/ step pulse request latched
        fPosNow_um := fPosNow_um + fDirSign * fEquivUse;   // 位置 LREAL 累加 [微米]（含方向符号）/ position accumulated with direction
    END_WHILE
    // 运动中越限急停：位置一旦离开软限位区间立即拦截 / in-motion overtravel e-stop
    IF (fPosNow_um > fUpUse + DL_STZ_TOL) OR (fPosNow_um < fLoUse - DL_STZ_TOL) THEN
        eState := E_DL_StepZState.eFault;             // 急停进故障态 / e-stop to fault
        eErr := E_DL_StepZErr.eLimitHit;              // 故障级：限位拦截 / fault: limit hit
        bLimitHit := TRUE;                            // 限位标志锁存 / limit flag latched
        bMoving := FALSE;                             // 运动撤 / moving dropped
        bStepPulse := FALSE;                          // 脉冲撤 / pulse dropped
        bStepReq := FALSE;                            // 脉冲请求撤 / pulse request dropped
        nStepsDone := nStepsTotal;                    // 终止本程 / terminate the move
    ELSIF nStepsDone >= nStepsTotal THEN
        eState := E_DL_StepZState.eDone;              // 步数发完：到位 / steps done: in position
        eErr := E_DL_StepZErr.eInPos;                 // 到位码 / in-position code
        bMoving := FALSE;                             // 运动撤 / moving dropped
    END_IF
END_IF

(*------------------------------------------------------------------------------
 * 段 7｜状态码映射与 CASE 兜底
 *----------------------------------------------------------------------------*)
CASE eState OF
    E_DL_StepZState.eIdle:
        IF (eErr <> E_DL_StepZErr.eConfigBad) AND (eErr <> E_DL_StepZErr.eTargetBad) AND (eErr <> E_DL_StepZErr.eLimitHit) THEN
            eErr := E_DL_StepZErr.eReady;             // 无挂起故障时保持就绪码 / ready code unless a fault is pending
        END_IF
    E_DL_StepZState.eMoving:
        bMoving := TRUE;                              // 运动相运动标志保持 / moving flag held in motion phase
    E_DL_StepZState.eDone:
        eErr := E_DL_StepZErr.eInPos;                 // 到位码 / in-position code
    E_DL_StepZState.eFault:
        bMoving := FALSE;                             // 故障态运动撤 / moving dropped in fault
        bStepPulse := FALSE;                          // 故障态脉冲撤 / pulse dropped in fault
        bStepReq := FALSE;                            // 故障态请求撤 / request dropped in fault
    ELSE
        eState := E_DL_StepZState.eFault;             // 非法状态兜底 / illegal-state fallback
        eErr := E_DL_StepZErr.eConfigBad;             // 兜底码（配置段，反证句：输出同为运动撤+故障级）/ fallback code
        bMoving := FALSE;                             // 运动撤 / moving dropped
        bStepPulse := FALSE;                          // 脉冲撤 / pulse dropped
        bStepReq := FALSE;                            // 请求撤 / request dropped
END_CASE
END_FUNCTION_BLOCK
